(* IEC 61131-3 sources: 2026_Projet_YGO_ExcavatriceDragage/TOOLS/TEST_AUTO_CI/RESULTS/L_SIMULATION/tests (part 2) *)

TEST 'TC-T418-005 Perte permis stimulus et conflit en mouvement'
VAR
    fb : FB_Sim_Joystick;
    i : INT;
END_VAR
    fb.Enable := TRUE; fb(); fb.BtnRev_Down_Open := TRUE;
    ADVANCE_TIME(10000000); fb();
ADVANCE_TIME(10000000); fb();
ADVANCE_TIME(10000000); fb();
ADVANCE_TIME(10000000); fb();
ADVANCE_TIME(10000000); fb();
ADVANCE_TIME(10000000); fb();
ADVANCE_TIME(10000000); fb();
ADVANCE_TIME(10000000); fb();
ADVANCE_TIME(10000000); fb();
ADVANCE_TIME(10000000); fb();
ADVANCE_TIME(10000000); fb();
ADVANCE_TIME(10000000); fb();
ADVANCE_TIME(10000000); fb();
ADVANCE_TIME(10000000); fb();
ADVANCE_TIME(10000000); fb();
ADVANCE_TIME(10000000); fb();
ADVANCE_TIME(10000000); fb();
ADVANCE_TIME(10000000); fb();
ADVANCE_TIME(10000000); fb();
ADVANCE_TIME(10000000); fb();
ADVANCE_TIME(10000000); fb();
ADVANCE_TIME(10000000); fb();
ADVANCE_TIME(10000000); fb();
ADVANCE_TIME(10000000); fb();
ADVANCE_TIME(10000000); fb();
ADVANCE_TIME(10000000); fb();
ADVANCE_TIME(10000000); fb();
ADVANCE_TIME(10000000); fb();
ADVANCE_TIME(10000000); fb();
ADVANCE_TIME(10000000); fb();
ADVANCE_TIME(10000000); fb();
ADVANCE_TIME(10000000); fb();
ADVANCE_TIME(10000000); fb();
ADVANCE_TIME(10000000); fb();
ADVANCE_TIME(10000000); fb();
ADVANCE_TIME(10000000); fb();
ADVANCE_TIME(10000000); fb();
ADVANCE_TIME(10000000); fb();
ADVANCE_TIME(10000000); fb();
ADVANCE_TIME(10000000); fb();
ADVANCE_TIME(10000000); fb();
ADVANCE_TIME(10000000); fb();
ADVANCE_TIME(10000000); fb();
ADVANCE_TIME(10000000); fb();
ADVANCE_TIME(10000000); fb();
ADVANCE_TIME(10000000); fb();
ADVANCE_TIME(10000000); fb();
ADVANCE_TIME(10000000); fb();
ADVANCE_TIME(10000000); fb();
ADVANCE_TIME(10000000); fb();
ADVANCE_TIME(10000000); fb();
ADVANCE_TIME(10000000); fb();
ADVANCE_TIME(10000000); fb();
ADVANCE_TIME(10000000); fb();
ADVANCE_TIME(10000000); fb();
ADVANCE_TIME(10000000); fb();
ADVANCE_TIME(10000000); fb();
ADVANCE_TIME(10000000); fb();
ADVANCE_TIME(10000000); fb();
ADVANCE_TIME(10000000); fb();
ADVANCE_TIME(10000000); fb();
ADVANCE_TIME(10000000); fb();
ADVANCE_TIME(10000000); fb();
ADVANCE_TIME(10000000); fb();
ADVANCE_TIME(10000000); fb();
ADVANCE_TIME(10000000); fb();
ADVANCE_TIME(10000000); fb();
ADVANCE_TIME(10000000); fb();
ADVANCE_TIME(10000000); fb();
ADVANCE_TIME(10000000); fb();
ADVANCE_TIME(10000000); fb();
ADVANCE_TIME(10000000); fb();
ADVANCE_TIME(10000000); fb();
ADVANCE_TIME(10000000); fb();
ADVANCE_TIME(10000000); fb();
ADVANCE_TIME(10000000); fb();
ADVANCE_TIME(10000000); fb();
ADVANCE_TIME(10000000); fb();
ADVANCE_TIME(10000000); fb();
ADVANCE_TIME(10000000); fb();
ADVANCE_TIME(10000000); fb();
ADVANCE_TIME(10000000); fb();
ADVANCE_TIME(10000000); fb();
ADVANCE_TIME(10000000); fb();
ADVANCE_TIME(10000000); fb();
ADVANCE_TIME(10000000); fb();
ADVANCE_TIME(10000000); fb();
ADVANCE_TIME(10000000); fb();
ADVANCE_TIME(10000000); fb();
ADVANCE_TIME(10000000); fb();
ADVANCE_TIME(10000000); fb();
ADVANCE_TIME(10000000); fb();
ADVANCE_TIME(10000000); fb();
ADVANCE_TIME(10000000); fb();
ADVANCE_TIME(10000000); fb();
ADVANCE_TIME(10000000); fb();
ADVANCE_TIME(10000000); fb();
ADVANCE_TIME(10000000); fb();
ADVANCE_TIME(10000000); fb();
ADVANCE_TIME(10000000); fb();
    ASSERT_TRUE(fb.RawY < 5000, 'Y negatif');
    fb.GesturePermit := FALSE; fb();
    ASSERT_FALSE(fb.RawButton, 'Retrait permis simulateur annule bouton');
    fb.GesturePermit := TRUE;
    ADVANCE_TIME(10000000); fb();
        ASSERT_FALSE(fb.RawButton, 'Retour permis ne rearme pas');
ADVANCE_TIME(10000000); fb();
        ASSERT_FALSE(fb.RawButton, 'Retour permis ne rearme pas');
ADVANCE_TIME(10000000); fb();
        ASSERT_FALSE(fb.RawButton, 'Retour permis ne rearme pas');
ADVANCE_TIME(10000000); fb();
        ASSERT_FALSE(fb.RawButton, 'Retour permis ne rearme pas');
ADVANCE_TIME(10000000); fb();
        ASSERT_FALSE(fb.RawButton, 'Retour permis ne rearme pas');
ADVANCE_TIME(10000000); fb();
        ASSERT_FALSE(fb.RawButton, 'Retour permis ne rearme pas');
ADVANCE_TIME(10000000); fb();
        ASSERT_FALSE(fb.RawButton, 'Retour permis ne rearme pas');
ADVANCE_TIME(10000000); fb();
        ASSERT_FALSE(fb.RawButton, 'Retour permis ne rearme pas');
ADVANCE_TIME(10000000); fb();
        ASSERT_FALSE(fb.RawButton, 'Retour permis ne rearme pas');
ADVANCE_TIME(10000000); fb();
        ASSERT_FALSE(fb.RawButton, 'Retour permis ne rearme pas');
ADVANCE_TIME(10000000); fb();
        ASSERT_FALSE(fb.RawButton, 'Retour permis ne rearme pas');
ADVANCE_TIME(10000000); fb();
        ASSERT_FALSE(fb.RawButton, 'Retour permis ne rearme pas');
ADVANCE_TIME(10000000); fb();
        ASSERT_FALSE(fb.RawButton, 'Retour permis ne rearme pas');
ADVANCE_TIME(10000000); fb();
        ASSERT_FALSE(fb.RawButton, 'Retour permis ne rearme pas');
ADVANCE_TIME(10000000); fb();
        ASSERT_FALSE(fb.RawButton, 'Retour permis ne rearme pas');
ADVANCE_TIME(10000000); fb();
        ASSERT_FALSE(fb.RawButton, 'Retour permis ne rearme pas');
ADVANCE_TIME(10000000); fb();
        ASSERT_FALSE(fb.RawButton, 'Retour permis ne rearme pas');
ADVANCE_TIME(10000000); fb();
        ASSERT_FALSE(fb.RawButton, 'Retour permis ne rearme pas');
ADVANCE_TIME(10000000); fb();
        ASSERT_FALSE(fb.RawButton, 'Retour permis ne rearme pas');
ADVANCE_TIME(10000000); fb();
        ASSERT_FALSE(fb.RawButton, 'Retour permis ne rearme pas');
ADVANCE_TIME(10000000); fb();
        ASSERT_FALSE(fb.RawButton, 'Retour permis ne rearme pas');
ADVANCE_TIME(10000000); fb();
        ASSERT_FALSE(fb.RawButton, 'Retour permis ne rearme pas');
ADVANCE_TIME(10000000); fb();
        ASSERT_FALSE(fb.RawButton, 'Retour permis ne rearme pas');
ADVANCE_TIME(10000000); fb();
        ASSERT_FALSE(fb.RawButton, 'Retour permis ne rearme pas');
ADVANCE_TIME(10000000); fb();
        ASSERT_FALSE(fb.RawButton, 'Retour permis ne rearme pas');
ADVANCE_TIME(10000000); fb();
        ASSERT_FALSE(fb.RawButton, 'Retour permis ne rearme pas');
ADVANCE_TIME(10000000); fb();
        ASSERT_FALSE(fb.RawButton, 'Retour permis ne rearme pas');
ADVANCE_TIME(10000000); fb();
        ASSERT_FALSE(fb.RawButton, 'Retour permis ne rearme pas');
ADVANCE_TIME(10000000); fb();
        ASSERT_FALSE(fb.RawButton, 'Retour permis ne rearme pas');
ADVANCE_TIME(10000000); fb();
        ASSERT_FALSE(fb.RawButton, 'Retour permis ne rearme pas');
ADVANCE_TIME(10000000); fb();
        ASSERT_FALSE(fb.RawButton, 'Retour permis ne rearme pas');
ADVANCE_TIME(10000000); fb();
        ASSERT_FALSE(fb.RawButton, 'Retour permis ne rearme pas');
ADVANCE_TIME(10000000); fb();
        ASSERT_FALSE(fb.RawButton, 'Retour permis ne rearme pas');
ADVANCE_TIME(10000000); fb();
        ASSERT_FALSE(fb.RawButton, 'Retour permis ne rearme pas');
ADVANCE_TIME(10000000); fb();
        ASSERT_FALSE(fb.RawButton, 'Retour permis ne rearme pas');
ADVANCE_TIME(10000000); fb();
        ASSERT_FALSE(fb.RawButton, 'Retour permis ne rearme pas');
ADVANCE_TIME(10000000); fb();
        ASSERT_FALSE(fb.RawButton, 'Retour permis ne rearme pas');
ADVANCE_TIME(10000000); fb();
        ASSERT_FALSE(fb.RawButton, 'Retour permis ne rearme pas');
ADVANCE_TIME(10000000); fb();
        ASSERT_FALSE(fb.RawButton, 'Retour permis ne rearme pas');
ADVANCE_TIME(10000000); fb();
        ASSERT_FALSE(fb.RawButton, 'Retour permis ne rearme pas');
ADVANCE_TIME(10000000); fb();
        ASSERT_FALSE(fb.RawButton, 'Retour permis ne rearme pas');
ADVANCE_TIME(10000000); fb();
        ASSERT_FALSE(fb.RawButton, 'Retour permis ne rearme pas');
ADVANCE_TIME(10000000); fb();
        ASSERT_FALSE(fb.RawButton, 'Retour permis ne rearme pas');
ADVANCE_TIME(10000000); fb();
        ASSERT_FALSE(fb.RawButton, 'Retour permis ne rearme pas');
ADVANCE_TIME(10000000); fb();
        ASSERT_FALSE(fb.RawButton, 'Retour permis ne rearme pas');
ADVANCE_TIME(10000000); fb();
        ASSERT_FALSE(fb.RawButton, 'Retour permis ne rearme pas');
ADVANCE_TIME(10000000); fb();
        ASSERT_FALSE(fb.RawButton, 'Retour permis ne rearme pas');
ADVANCE_TIME(10000000); fb();
        ASSERT_FALSE(fb.RawButton, 'Retour permis ne rearme pas');
ADVANCE_TIME(10000000); fb();
        ASSERT_FALSE(fb.RawButton, 'Retour permis ne rearme pas');
ADVANCE_TIME(10000000); fb();
        ASSERT_FALSE(fb.RawButton, 'Retour permis ne rearme pas');
ADVANCE_TIME(10000000); fb();
        ASSERT_FALSE(fb.RawButton, 'Retour permis ne rearme pas');
ADVANCE_TIME(10000000); fb();
        ASSERT_FALSE(fb.RawButton, 'Retour permis ne rearme pas');
ADVANCE_TIME(10000000); fb();
        ASSERT_FALSE(fb.RawButton, 'Retour permis ne rearme pas');
ADVANCE_TIME(10000000); fb();
        ASSERT_FALSE(fb.RawButton, 'Retour permis ne rearme pas');
ADVANCE_TIME(10000000); fb();
        ASSERT_FALSE(fb.RawButton, 'Retour permis ne rearme pas');
ADVANCE_TIME(10000000); fb();
        ASSERT_FALSE(fb.RawButton, 'Retour permis ne rearme pas');
ADVANCE_TIME(10000000); fb();
        ASSERT_FALSE(fb.RawButton, 'Retour permis ne rearme pas');
ADVANCE_TIME(10000000); fb();
        ASSERT_FALSE(fb.RawButton, 'Retour permis ne rearme pas');
ADVANCE_TIME(10000000); fb();
        ASSERT_FALSE(fb.RawButton, 'Retour permis ne rearme pas');
ADVANCE_TIME(10000000); fb();
        ASSERT_FALSE(fb.RawButton, 'Retour permis ne rearme pas');
ADVANCE_TIME(10000000); fb();
        ASSERT_FALSE(fb.RawButton, 'Retour permis ne rearme pas');
ADVANCE_TIME(10000000); fb();
        ASSERT_FALSE(fb.RawButton, 'Retour permis ne rearme pas');
ADVANCE_TIME(10000000); fb();
        ASSERT_FALSE(fb.RawButton, 'Retour permis ne rearme pas');
ADVANCE_TIME(10000000); fb();
        ASSERT_FALSE(fb.RawButton, 'Retour permis ne rearme pas');
ADVANCE_TIME(10000000); fb();
        ASSERT_FALSE(fb.RawButton, 'Retour permis ne rearme pas');
ADVANCE_TIME(10000000); fb();
        ASSERT_FALSE(fb.RawButton, 'Retour permis ne rearme pas');
ADVANCE_TIME(10000000); fb();
        ASSERT_FALSE(fb.RawButton, 'Retour permis ne rearme pas');
ADVANCE_TIME(10000000); fb();
        ASSERT_FALSE(fb.RawButton, 'Retour permis ne rearme pas');
ADVANCE_TIME(10000000); fb();
        ASSERT_FALSE(fb.RawButton, 'Retour permis ne rearme pas');
ADVANCE_TIME(10000000); fb();
        ASSERT_FALSE(fb.RawButton, 'Retour permis ne rearme pas');
ADVANCE_TIME(10000000); fb();
        ASSERT_FALSE(fb.RawButton, 'Retour permis ne rearme pas');
ADVANCE_TIME(10000000); fb();
        ASSERT_FALSE(fb.RawButton, 'Retour permis ne rearme pas');
ADVANCE_TIME(10000000); fb();
        ASSERT_FALSE(fb.RawButton, 'Retour permis ne rearme pas');
ADVANCE_TIME(10000000); fb();
        ASSERT_FALSE(fb.RawButton, 'Retour permis ne rearme pas');
ADVANCE_TIME(10000000); fb();
        ASSERT_FALSE(fb.RawButton, 'Retour permis ne rearme pas');
ADVANCE_TIME(10000000); fb();
        ASSERT_FALSE(fb.RawButton, 'Retour permis ne rearme pas');
ADVANCE_TIME(10000000); fb();
        ASSERT_FALSE(fb.RawButton, 'Retour permis ne rearme pas');
ADVANCE_TIME(10000000); fb();
        ASSERT_FALSE(fb.RawButton, 'Retour permis ne rearme pas');
ADVANCE_TIME(10000000); fb();
        ASSERT_FALSE(fb.RawButton, 'Retour permis ne rearme pas');
ADVANCE_TIME(10000000); fb();
        ASSERT_FALSE(fb.RawButton, 'Retour permis ne rearme pas');
ADVANCE_TIME(10000000); fb();
        ASSERT_FALSE(fb.RawButton, 'Retour permis ne rearme pas');
ADVANCE_TIME(10000000); fb();
        ASSERT_FALSE(fb.RawButton, 'Retour permis ne rearme pas');
ADVANCE_TIME(10000000); fb();
        ASSERT_FALSE(fb.RawButton, 'Retour permis ne rearme pas');
ADVANCE_TIME(10000000); fb();
        ASSERT_FALSE(fb.RawButton, 'Retour permis ne rearme pas');
ADVANCE_TIME(10000000); fb();
        ASSERT_FALSE(fb.RawButton, 'Retour permis ne rearme pas');
ADVANCE_TIME(10000000); fb();
        ASSERT_FALSE(fb.RawButton, 'Retour permis ne rearme pas');
ADVANCE_TIME(10000000); fb();
        ASSERT_FALSE(fb.RawButton, 'Retour permis ne rearme pas');
ADVANCE_TIME(10000000); fb();
        ASSERT_FALSE(fb.RawButton, 'Retour permis ne rearme pas');
ADVANCE_TIME(10000000); fb();
        ASSERT_FALSE(fb.RawButton, 'Retour permis ne rearme pas');
ADVANCE_TIME(10000000); fb();
        ASSERT_FALSE(fb.RawButton, 'Retour permis ne rearme pas');
ADVANCE_TIME(10000000); fb();
        ASSERT_FALSE(fb.RawButton, 'Retour permis ne rearme pas');
ADVANCE_TIME(10000000); fb();
        ASSERT_FALSE(fb.RawButton, 'Retour permis ne rearme pas');
ADVANCE_TIME(10000000); fb();
        ASSERT_FALSE(fb.RawButton, 'Retour permis ne rearme pas');
ADVANCE_TIME(10000000); fb();
        ASSERT_FALSE(fb.RawButton, 'Retour permis ne rearme pas');
ADVANCE_TIME(10000000); fb();
        ASSERT_FALSE(fb.RawButton, 'Retour permis ne rearme pas');
ADVANCE_TIME(10000000); fb();
        ASSERT_FALSE(fb.RawButton, 'Retour permis ne rearme pas');
ADVANCE_TIME(10000000); fb();
        ASSERT_FALSE(fb.RawButton, 'Retour permis ne rearme pas');
ADVANCE_TIME(10000000); fb();
        ASSERT_FALSE(fb.RawButton, 'Retour permis ne rearme pas');
ADVANCE_TIME(10000000); fb();
        ASSERT_FALSE(fb.RawButton, 'Retour permis ne rearme pas');
ADVANCE_TIME(10000000); fb();
        ASSERT_FALSE(fb.RawButton, 'Retour permis ne rearme pas');
    ASSERT_EQ(fb.RawY, 5000, 'Retour neutre');
    fb.BtnRev_Down_Open := FALSE; fb(); fb.BtnFwd_Up_Close := TRUE;
    ADVANCE_TIME(10000000); fb();
ADVANCE_TIME(10000000); fb();
ADVANCE_TIME(10000000); fb();
ADVANCE_TIME(10000000); fb();
ADVANCE_TIME(10000000); fb();
ADVANCE_TIME(10000000); fb();
ADVANCE_TIME(10000000); fb();
ADVANCE_TIME(10000000); fb();
ADVANCE_TIME(10000000); fb();
ADVANCE_TIME(10000000); fb();
ADVANCE_TIME(10000000); fb();
ADVANCE_TIME(10000000); fb();
ADVANCE_TIME(10000000); fb();
ADVANCE_TIME(10000000); fb();
ADVANCE_TIME(10000000); fb();
ADVANCE_TIME(10000000); fb();
ADVANCE_TIME(10000000); fb();
ADVANCE_TIME(10000000); fb();
ADVANCE_TIME(10000000); fb();
ADVANCE_TIME(10000000); fb();
ADVANCE_TIME(10000000); fb();
ADVANCE_TIME(10000000); fb();
ADVANCE_TIME(10000000); fb();
ADVANCE_TIME(10000000); fb();
ADVANCE_TIME(10000000); fb();
ADVANCE_TIME(10000000); fb();
ADVANCE_TIME(10000000); fb();
ADVANCE_TIME(10000000); fb();
ADVANCE_TIME(10000000); fb();
ADVANCE_TIME(10000000); fb();
ADVANCE_TIME(10000000); fb();
ADVANCE_TIME(10000000); fb();
ADVANCE_TIME(10000000); fb();
ADVANCE_TIME(10000000); fb();
ADVANCE_TIME(10000000); fb();
ADVANCE_TIME(10000000); fb();
ADVANCE_TIME(10000000); fb();
ADVANCE_TIME(10000000); fb();
ADVANCE_TIME(10000000); fb();
ADVANCE_TIME(10000000); fb();
ADVANCE_TIME(10000000); fb();
ADVANCE_TIME(10000000); fb();
ADVANCE_TIME(10000000); fb();
ADVANCE_TIME(10000000); fb();
ADVANCE_TIME(10000000); fb();
ADVANCE_TIME(10000000); fb();
ADVANCE_TIME(10000000); fb();
ADVANCE_TIME(10000000); fb();
ADVANCE_TIME(10000000); fb();
ADVANCE_TIME(10000000); fb();
ADVANCE_TIME(10000000); fb();
ADVANCE_TIME(10000000); fb();
ADVANCE_TIME(10000000); fb();
ADVANCE_TIME(10000000); fb();
ADVANCE_TIME(10000000); fb();
ADVANCE_TIME(10000000); fb();
ADVANCE_TIME(10000000); fb();
ADVANCE_TIME(10000000); fb();
ADVANCE_TIME(10000000); fb();
ADVANCE_TIME(10000000); fb();
ADVANCE_TIME(10000000); fb();
ADVANCE_TIME(10000000); fb();
ADVANCE_TIME(10000000); fb();
ADVANCE_TIME(10000000); fb();
ADVANCE_TIME(10000000); fb();
ADVANCE_TIME(10000000); fb();
ADVANCE_TIME(10000000); fb();
ADVANCE_TIME(10000000); fb();
ADVANCE_TIME(10000000); fb();
ADVANCE_TIME(10000000); fb();
ADVANCE_TIME(10000000); fb();
ADVANCE_TIME(10000000); fb();
ADVANCE_TIME(10000000); fb();
ADVANCE_TIME(10000000); fb();
ADVANCE_TIME(10000000); fb();
ADVANCE_TIME(10000000); fb();
ADVANCE_TIME(10000000); fb();
ADVANCE_TIME(10000000); fb();
ADVANCE_TIME(10000000); fb();
ADVANCE_TIME(10000000); fb();
ADVANCE_TIME(10000000); fb();
ADVANCE_TIME(10000000); fb();
ADVANCE_TIME(10000000); fb();
ADVANCE_TIME(10000000); fb();
ADVANCE_TIME(10000000); fb();
ADVANCE_TIME(10000000); fb();
ADVANCE_TIME(10000000); fb();
ADVANCE_TIME(10000000); fb();
ADVANCE_TIME(10000000); fb();
ADVANCE_TIME(10000000); fb();
ADVANCE_TIME(10000000); fb();
ADVANCE_TIME(10000000); fb();
ADVANCE_TIME(10000000); fb();
ADVANCE_TIME(10000000); fb();
ADVANCE_TIME(10000000); fb();
ADVANCE_TIME(10000000); fb();
ADVANCE_TIME(10000000); fb();
ADVANCE_TIME(10000000); fb();
ADVANCE_TIME(10000000); fb();
ADVANCE_TIME(10000000); fb();
    fb.BtnRight_Fwd_MAINT := TRUE;
    ADVANCE_TIME(10000000); fb();
ADVANCE_TIME(10000000); fb();
ADVANCE_TIME(10000000); fb();
ADVANCE_TIME(10000000); fb();
ADVANCE_TIME(10000000); fb();
ADVANCE_TIME(10000000); fb();
ADVANCE_TIME(10000000); fb();
ADVANCE_TIME(10000000); fb();
ADVANCE_TIME(10000000); fb();
ADVANCE_TIME(10000000); fb();
ADVANCE_TIME(10000000); fb();
ADVANCE_TIME(10000000); fb();
ADVANCE_TIME(10000000); fb();
ADVANCE_TIME(10000000); fb();
ADVANCE_TIME(10000000); fb();
ADVANCE_TIME(10000000); fb();
ADVANCE_TIME(10000000); fb();
ADVANCE_TIME(10000000); fb();
ADVANCE_TIME(10000000); fb();
ADVANCE_TIME(10000000); fb();
ADVANCE_TIME(10000000); fb();
ADVANCE_TIME(10000000); fb();
ADVANCE_TIME(10000000); fb();
ADVANCE_TIME(10000000); fb();
ADVANCE_TIME(10000000); fb();
ADVANCE_TIME(10000000); fb();
ADVANCE_TIME(10000000); fb();
ADVANCE_TIME(10000000); fb();
ADVANCE_TIME(10000000); fb();
ADVANCE_TIME(10000000); fb();
ADVANCE_TIME(10000000); fb();
ADVANCE_TIME(10000000); fb();
ADVANCE_TIME(10000000); fb();
ADVANCE_TIME(10000000); fb();
ADVANCE_TIME(10000000); fb();
ADVANCE_TIME(10000000); fb();
ADVANCE_TIME(10000000); fb();
ADVANCE_TIME(10000000); fb();
ADVANCE_TIME(10000000); fb();
ADVANCE_TIME(10000000); fb();
ADVANCE_TIME(10000000); fb();
ADVANCE_TIME(10000000); fb();
ADVANCE_TIME(10000000); fb();
ADVANCE_TIME(10000000); fb();
ADVANCE_TIME(10000000); fb();
ADVANCE_TIME(10000000); fb();
ADVANCE_TIME(10000000); fb();
ADVANCE_TIME(10000000); fb();
ADVANCE_TIME(10000000); fb();
ADVANCE_TIME(10000000); fb();
ADVANCE_TIME(10000000); fb();
ADVANCE_TIME(10000000); fb();
ADVANCE_TIME(10000000); fb();
ADVANCE_TIME(10000000); fb();
ADVANCE_TIME(10000000); fb();
ADVANCE_TIME(10000000); fb();
ADVANCE_TIME(10000000); fb();
ADVANCE_TIME(10000000); fb();
ADVANCE_TIME(10000000); fb();
ADVANCE_TIME(10000000); fb();
ADVANCE_TIME(10000000); fb();
ADVANCE_TIME(10000000); fb();
ADVANCE_TIME(10000000); fb();
ADVANCE_TIME(10000000); fb();
ADVANCE_TIME(10000000); fb();
ADVANCE_TIME(10000000); fb();
ADVANCE_TIME(10000000); fb();
ADVANCE_TIME(10000000); fb();
ADVANCE_TIME(10000000); fb();
ADVANCE_TIME(10000000); fb();
ADVANCE_TIME(10000000); fb();
ADVANCE_TIME(10000000); fb();
ADVANCE_TIME(10000000); fb();
ADVANCE_TIME(10000000); fb();
ADVANCE_TIME(10000000); fb();
ADVANCE_TIME(10000000); fb();
ADVANCE_TIME(10000000); fb();
ADVANCE_TIME(10000000); fb();
ADVANCE_TIME(10000000); fb();
ADVANCE_TIME(10000000); fb();
ADVANCE_TIME(10000000); fb();
ADVANCE_TIME(10000000); fb();
ADVANCE_TIME(10000000); fb();
ADVANCE_TIME(10000000); fb();
ADVANCE_TIME(10000000); fb();
ADVANCE_TIME(10000000); fb();
ADVANCE_TIME(10000000); fb();
ADVANCE_TIME(10000000); fb();
ADVANCE_TIME(10000000); fb();
ADVANCE_TIME(10000000); fb();
ADVANCE_TIME(10000000); fb();
ADVANCE_TIME(10000000); fb();
ADVANCE_TIME(10000000); fb();
ADVANCE_TIME(10000000); fb();
ADVANCE_TIME(10000000); fb();
ADVANCE_TIME(10000000); fb();
ADVANCE_TIME(10000000); fb();
ADVANCE_TIME(10000000); fb();
ADVANCE_TIME(10000000); fb();
ADVANCE_TIME(10000000); fb();
    ASSERT_EQ(fb.RawY, 5000, 'Conflit en mouvement retourne au neutre');
    ASSERT_FALSE(fb.RawButton, 'Conflit ne produit pas appui');
END_TEST

TEST 'TC-T418-006 Dynamiques depassement et bagotement conservees'
VAR
    fb : FB_Sim_Joystick;
    i : INT;
    oscillationSeen : BOOL;
END_VAR
    oscillationSeen := FALSE;
    fb.Enable := TRUE; fb.OvershootActive := TRUE; fb.BagotementActive := TRUE;
    fb(); fb.BtnRight_Fwd_MAINT := TRUE;
    ADVANCE_TIME(10000000); fb();
ADVANCE_TIME(10000000); fb();
ADVANCE_TIME(10000000); fb();
ADVANCE_TIME(10000000); fb();
ADVANCE_TIME(10000000); fb();
ADVANCE_TIME(10000000); fb();
ADVANCE_TIME(10000000); fb();
ADVANCE_TIME(10000000); fb();
ADVANCE_TIME(10000000); fb();
ADVANCE_TIME(10000000); fb();
ADVANCE_TIME(10000000); fb();
ADVANCE_TIME(10000000); fb();
ADVANCE_TIME(10000000); fb();
ADVANCE_TIME(10000000); fb();
ADVANCE_TIME(10000000); fb();
ADVANCE_TIME(10000000); fb();
ADVANCE_TIME(10000000); fb();
ADVANCE_TIME(10000000); fb();
ADVANCE_TIME(10000000); fb();
ADVANCE_TIME(10000000); fb();
ADVANCE_TIME(10000000); fb();
ADVANCE_TIME(10000000); fb();
ADVANCE_TIME(10000000); fb();
ADVANCE_TIME(10000000); fb();
ADVANCE_TIME(10000000); fb();
ADVANCE_TIME(10000000); fb();
ADVANCE_TIME(10000000); fb();
ADVANCE_TIME(10000000); fb();
ADVANCE_TIME(10000000); fb();
ADVANCE_TIME(10000000); fb();
ADVANCE_TIME(10000000); fb();
ADVANCE_TIME(10000000); fb();
ADVANCE_TIME(10000000); fb();
ADVANCE_TIME(10000000); fb();
ADVANCE_TIME(10000000); fb();
ADVANCE_TIME(10000000); fb();
ADVANCE_TIME(10000000); fb();
ADVANCE_TIME(10000000); fb();
ADVANCE_TIME(10000000); fb();
ADVANCE_TIME(10000000); fb();
ADVANCE_TIME(10000000); fb();
ADVANCE_TIME(10000000); fb();
ADVANCE_TIME(10000000); fb();
ADVANCE_TIME(10000000); fb();
ADVANCE_TIME(10000000); fb();
ADVANCE_TIME(10000000); fb();
ADVANCE_TIME(10000000); fb();
ADVANCE_TIME(10000000); fb();
ADVANCE_TIME(10000000); fb();
ADVANCE_TIME(10000000); fb();
ADVANCE_TIME(10000000); fb();
ADVANCE_TIME(10000000); fb();
ADVANCE_TIME(10000000); fb();
ADVANCE_TIME(10000000); fb();
ADVANCE_TIME(10000000); fb();
ADVANCE_TIME(10000000); fb();
ADVANCE_TIME(10000000); fb();
ADVANCE_TIME(10000000); fb();
ADVANCE_TIME(10000000); fb();
ADVANCE_TIME(10000000); fb();
ADVANCE_TIME(10000000); fb();
ADVANCE_TIME(10000000); fb();
ADVANCE_TIME(10000000); fb();
ADVANCE_TIME(10000000); fb();
ADVANCE_TIME(10000000); fb();
ADVANCE_TIME(10000000); fb();
ADVANCE_TIME(10000000); fb();
ADVANCE_TIME(10000000); fb();
ADVANCE_TIME(10000000); fb();
ADVANCE_TIME(10000000); fb();
ADVANCE_TIME(10000000); fb();
ADVANCE_TIME(10000000); fb();
ADVANCE_TIME(10000000); fb();
ADVANCE_TIME(10000000); fb();
ADVANCE_TIME(10000000); fb();
ADVANCE_TIME(10000000); fb();
ADVANCE_TIME(10000000); fb();
ADVANCE_TIME(10000000); fb();
ADVANCE_TIME(10000000); fb();
ADVANCE_TIME(10000000); fb();
ADVANCE_TIME(10000000); fb();
ADVANCE_TIME(10000000); fb();
ADVANCE_TIME(10000000); fb();
ADVANCE_TIME(10000000); fb();
ADVANCE_TIME(10000000); fb();
ADVANCE_TIME(10000000); fb();
ADVANCE_TIME(10000000); fb();
ADVANCE_TIME(10000000); fb();
ADVANCE_TIME(10000000); fb();
ADVANCE_TIME(10000000); fb();
ADVANCE_TIME(10000000); fb();
ADVANCE_TIME(10000000); fb();
ADVANCE_TIME(10000000); fb();
ADVANCE_TIME(10000000); fb();
ADVANCE_TIME(10000000); fb();
ADVANCE_TIME(10000000); fb();
ADVANCE_TIME(10000000); fb();
ADVANCE_TIME(10000000); fb();
ADVANCE_TIME(10000000); fb();
ADVANCE_TIME(10000000); fb();
ADVANCE_TIME(10000000); fb();
ADVANCE_TIME(10000000); fb();
ADVANCE_TIME(10000000); fb();
ADVANCE_TIME(10000000); fb();
ADVANCE_TIME(10000000); fb();
ADVANCE_TIME(10000000); fb();
ADVANCE_TIME(10000000); fb();
ADVANCE_TIME(10000000); fb();
ADVANCE_TIME(10000000); fb();
ADVANCE_TIME(10000000); fb();
ADVANCE_TIME(10000000); fb();
ADVANCE_TIME(10000000); fb();
ADVANCE_TIME(10000000); fb();
ADVANCE_TIME(10000000); fb();
ADVANCE_TIME(10000000); fb();
ADVANCE_TIME(10000000); fb();
ADVANCE_TIME(10000000); fb();
ADVANCE_TIME(10000000); fb();
ADVANCE_TIME(10000000); fb();
ADVANCE_TIME(10000000); fb();
ADVANCE_TIME(10000000); fb();
ADVANCE_TIME(10000000); fb();
ADVANCE_TIME(10000000); fb();
ADVANCE_TIME(10000000); fb();
ADVANCE_TIME(10000000); fb();
ADVANCE_TIME(10000000); fb();
ADVANCE_TIME(10000000); fb();
ADVANCE_TIME(10000000); fb();
ADVANCE_TIME(10000000); fb();
ADVANCE_TIME(10000000); fb();
ADVANCE_TIME(10000000); fb();
ADVANCE_TIME(10000000); fb();
ADVANCE_TIME(10000000); fb();
ADVANCE_TIME(10000000); fb();
ADVANCE_TIME(10000000); fb();
ADVANCE_TIME(10000000); fb();
ADVANCE_TIME(10000000); fb();
ADVANCE_TIME(10000000); fb();
ADVANCE_TIME(10000000); fb();
ADVANCE_TIME(10000000); fb();
ADVANCE_TIME(10000000); fb();
ADVANCE_TIME(10000000); fb();
ADVANCE_TIME(10000000); fb();
ADVANCE_TIME(10000000); fb();
ADVANCE_TIME(10000000); fb();
ADVANCE_TIME(10000000); fb();
ADVANCE_TIME(10000000); fb();
ADVANCE_TIME(10000000); fb();
ADVANCE_TIME(10000000); fb();
ADVANCE_TIME(10000000); fb();
ADVANCE_TIME(10000000); fb();
ADVANCE_TIME(10000000); fb();
ADVANCE_TIME(10000000); fb();
ADVANCE_TIME(10000000); fb();
ADVANCE_TIME(10000000); fb();
ADVANCE_TIME(10000000); fb();
ADVANCE_TIME(10000000); fb();
ADVANCE_TIME(10000000); fb();
ADVANCE_TIME(10000000); fb();
ADVANCE_TIME(10000000); fb();
ADVANCE_TIME(10000000); fb();
ADVANCE_TIME(10000000); fb();
ADVANCE_TIME(10000000); fb();
ADVANCE_TIME(10000000); fb();
ADVANCE_TIME(10000000); fb();
ADVANCE_TIME(10000000); fb();
ADVANCE_TIME(10000000); fb();
ADVANCE_TIME(10000000); fb();
ADVANCE_TIME(10000000); fb();
ADVANCE_TIME(10000000); fb();
ADVANCE_TIME(10000000); fb();
ADVANCE_TIME(10000000); fb();
ADVANCE_TIME(10000000); fb();
ADVANCE_TIME(10000000); fb();
ADVANCE_TIME(10000000); fb();
ADVANCE_TIME(10000000); fb();
ADVANCE_TIME(10000000); fb();
ADVANCE_TIME(10000000); fb();
ADVANCE_TIME(10000000); fb();
ADVANCE_TIME(10000000); fb();
ADVANCE_TIME(10000000); fb();
ADVANCE_TIME(10000000); fb();
ADVANCE_TIME(10000000); fb();
ADVANCE_TIME(10000000); fb();
ADVANCE_TIME(10000000); fb();
ADVANCE_TIME(10000000); fb();
ADVANCE_TIME(10000000); fb();
ADVANCE_TIME(10000000); fb();
ADVANCE_TIME(10000000); fb();
ADVANCE_TIME(10000000); fb();
ADVANCE_TIME(10000000); fb();
ADVANCE_TIME(10000000); fb();
ADVANCE_TIME(10000000); fb();
ADVANCE_TIME(10000000); fb();
ADVANCE_TIME(10000000); fb();
ADVANCE_TIME(10000000); fb();
ADVANCE_TIME(10000000); fb();
ADVANCE_TIME(10000000); fb();
ADVANCE_TIME(10000000); fb();
ADVANCE_TIME(10000000); fb();
ADVANCE_TIME(10000000); fb();
ADVANCE_TIME(10000000); fb();
ADVANCE_TIME(10000000); fb();
ADVANCE_TIME(10000000); fb();
ADVANCE_TIME(10000000); fb();
ADVANCE_TIME(10000000); fb();
ADVANCE_TIME(10000000); fb();
ADVANCE_TIME(10000000); fb();
ADVANCE_TIME(10000000); fb();
ADVANCE_TIME(10000000); fb();
ADVANCE_TIME(10000000); fb();
ADVANCE_TIME(10000000); fb();
ADVANCE_TIME(10000000); fb();
ADVANCE_TIME(10000000); fb();
ADVANCE_TIME(10000000); fb();
ADVANCE_TIME(10000000); fb();
ADVANCE_TIME(10000000); fb();
ADVANCE_TIME(10000000); fb();
ADVANCE_TIME(10000000); fb();
ADVANCE_TIME(10000000); fb();
ADVANCE_TIME(10000000); fb();
ADVANCE_TIME(10000000); fb();
ADVANCE_TIME(10000000); fb();
ADVANCE_TIME(10000000); fb();
ADVANCE_TIME(10000000); fb();
ADVANCE_TIME(10000000); fb();
ADVANCE_TIME(10000000); fb();
ADVANCE_TIME(10000000); fb();
ADVANCE_TIME(10000000); fb();
ADVANCE_TIME(10000000); fb();
ADVANCE_TIME(10000000); fb();
ADVANCE_TIME(10000000); fb();
ADVANCE_TIME(10000000); fb();
ADVANCE_TIME(10000000); fb();
ADVANCE_TIME(10000000); fb();
ADVANCE_TIME(10000000); fb();
ADVANCE_TIME(10000000); fb();
ADVANCE_TIME(10000000); fb();
ADVANCE_TIME(10000000); fb();
ADVANCE_TIME(10000000); fb();
ADVANCE_TIME(10000000); fb();
ADVANCE_TIME(10000000); fb();
ADVANCE_TIME(10000000); fb();
ADVANCE_TIME(10000000); fb();
ADVANCE_TIME(10000000); fb();
ADVANCE_TIME(10000000); fb();
ADVANCE_TIME(10000000); fb();
ADVANCE_TIME(10000000); fb();
ADVANCE_TIME(10000000); fb();
ADVANCE_TIME(10000000); fb();
    ASSERT_TRUE(fb.RawX > 10500, 'Injection depassement capteur conservee');
    fb.BtnRight_Fwd_MAINT := FALSE;
    ADVANCE_TIME(10000000); fb();
        IF fb.RawX < 5000 THEN oscillationSeen := TRUE; END_IF;
        ASSERT_FALSE(fb.RawButton, 'Aucun front pendant bagotement');
ADVANCE_TIME(10000000); fb();
        IF fb.RawX < 5000 THEN oscillationSeen := TRUE; END_IF;
        ASSERT_FALSE(fb.RawButton, 'Aucun front pendant bagotement');
ADVANCE_TIME(10000000); fb();
        IF fb.RawX < 5000 THEN oscillationSeen := TRUE; END_IF;
        ASSERT_FALSE(fb.RawButton, 'Aucun front pendant bagotement');
ADVANCE_TIME(10000000); fb();
        IF fb.RawX < 5000 THEN oscillationSeen := TRUE; END_IF;
        ASSERT_FALSE(fb.RawButton, 'Aucun front pendant bagotement');
ADVANCE_TIME(10000000); fb();
        IF fb.RawX < 5000 THEN oscillationSeen := TRUE; END_IF;
        ASSERT_FALSE(fb.RawButton, 'Aucun front pendant bagotement');
ADVANCE_TIME(10000000); fb();
        IF fb.RawX < 5000 THEN oscillationSeen := TRUE; END_IF;
        ASSERT_FALSE(fb.RawButton, 'Aucun front pendant bagotement');
ADVANCE_TIME(10000000); fb();
        IF fb.RawX < 5000 THEN oscillationSeen := TRUE; END_IF;
        ASSERT_FALSE(fb.RawButton, 'Aucun front pendant bagotement');
ADVANCE_TIME(10000000); fb();
        IF fb.RawX < 5000 THEN oscillationSeen := TRUE; END_IF;
        ASSERT_FALSE(fb.RawButton, 'Aucun front pendant bagotement');
ADVANCE_TIME(10000000); fb();
        IF fb.RawX < 5000 THEN oscillationSeen := TRUE; END_IF;
        ASSERT_FALSE(fb.RawButton, 'Aucun front pendant bagotement');
ADVANCE_TIME(10000000); fb();
        IF fb.RawX < 5000 THEN oscillationSeen := TRUE; END_IF;
        ASSERT_FALSE(fb.RawButton, 'Aucun front pendant bagotement');
ADVANCE_TIME(10000000); fb();
        IF fb.RawX < 5000 THEN oscillationSeen := TRUE; END_IF;
        ASSERT_FALSE(fb.RawButton, 'Aucun front pendant bagotement');
ADVANCE_TIME(10000000); fb();
        IF fb.RawX < 5000 THEN oscillationSeen := TRUE; END_IF;
        ASSERT_FALSE(fb.RawButton, 'Aucun front pendant bagotement');
ADVANCE_TIME(10000000); fb();
        IF fb.RawX < 5000 THEN oscillationSeen := TRUE; END_IF;
        ASSERT_FALSE(fb.RawButton, 'Aucun front pendant bagotement');
ADVANCE_TIME(10000000); fb();
        IF fb.RawX < 5000 THEN oscillationSeen := TRUE; END_IF;
        ASSERT_FALSE(fb.RawButton, 'Aucun front pendant bagotement');
ADVANCE_TIME(10000000); fb();
        IF fb.RawX < 5000 THEN oscillationSeen := TRUE; END_IF;
        ASSERT_FALSE(fb.RawButton, 'Aucun front pendant bagotement');
ADVANCE_TIME(10000000); fb();
        IF fb.RawX < 5000 THEN oscillationSeen := TRUE; END_IF;
        ASSERT_FALSE(fb.RawButton, 'Aucun front pendant bagotement');
ADVANCE_TIME(10000000); fb();
        IF fb.RawX < 5000 THEN oscillationSeen := TRUE; END_IF;
        ASSERT_FALSE(fb.RawButton, 'Aucun front pendant bagotement');
ADVANCE_TIME(10000000); fb();
        IF fb.RawX < 5000 THEN oscillationSeen := TRUE; END_IF;
        ASSERT_FALSE(fb.RawButton, 'Aucun front pendant bagotement');
ADVANCE_TIME(10000000); fb();
        IF fb.RawX < 5000 THEN oscillationSeen := TRUE; END_IF;
        ASSERT_FALSE(fb.RawButton, 'Aucun front pendant bagotement');
ADVANCE_TIME(10000000); fb();
        IF fb.RawX < 5000 THEN oscillationSeen := TRUE; END_IF;
        ASSERT_FALSE(fb.RawButton, 'Aucun front pendant bagotement');
ADVANCE_TIME(10000000); fb();
        IF fb.RawX < 5000 THEN oscillationSeen := TRUE; END_IF;
        ASSERT_FALSE(fb.RawButton, 'Aucun front pendant bagotement');
ADVANCE_TIME(10000000); fb();
        IF fb.RawX < 5000 THEN oscillationSeen := TRUE; END_IF;
        ASSERT_FALSE(fb.RawButton, 'Aucun front pendant bagotement');
ADVANCE_TIME(10000000); fb();
        IF fb.RawX < 5000 THEN oscillationSeen := TRUE; END_IF;
        ASSERT_FALSE(fb.RawButton, 'Aucun front pendant bagotement');
ADVANCE_TIME(10000000); fb();
        IF fb.RawX < 5000 THEN oscillationSeen := TRUE; END_IF;
        ASSERT_FALSE(fb.RawButton, 'Aucun front pendant bagotement');
ADVANCE_TIME(10000000); fb();
        IF fb.RawX < 5000 THEN oscillationSeen := TRUE; END_IF;
        ASSERT_FALSE(fb.RawButton, 'Aucun front pendant bagotement');
ADVANCE_TIME(10000000); fb();
        IF fb.RawX < 5000 THEN oscillationSeen := TRUE; END_IF;
        ASSERT_FALSE(fb.RawButton, 'Aucun front pendant bagotement');
ADVANCE_TIME(10000000); fb();
        IF fb.RawX < 5000 THEN oscillationSeen := TRUE; END_IF;
        ASSERT_FALSE(fb.RawButton, 'Aucun front pendant bagotement');
ADVANCE_TIME(10000000); fb();
        IF fb.RawX < 5000 THEN oscillationSeen := TRUE; END_IF;
        ASSERT_FALSE(fb.RawButton, 'Aucun front pendant bagotement');
ADVANCE_TIME(10000000); fb();
        IF fb.RawX < 5000 THEN oscillationSeen := TRUE; END_IF;
        ASSERT_FALSE(fb.RawButton, 'Aucun front pendant bagotement');
ADVANCE_TIME(10000000); fb();
        IF fb.RawX < 5000 THEN oscillationSeen := TRUE; END_IF;
        ASSERT_FALSE(fb.RawButton, 'Aucun front pendant bagotement');
ADVANCE_TIME(10000000); fb();
        IF fb.RawX < 5000 THEN oscillationSeen := TRUE; END_IF;
        ASSERT_FALSE(fb.RawButton, 'Aucun front pendant bagotement');
ADVANCE_TIME(10000000); fb();
        IF fb.RawX < 5000 THEN oscillationSeen := TRUE; END_IF;
        ASSERT_FALSE(fb.RawButton, 'Aucun front pendant bagotement');
ADVANCE_TIME(10000000); fb();
        IF fb.RawX < 5000 THEN oscillationSeen := TRUE; END_IF;
        ASSERT_FALSE(fb.RawButton, 'Aucun front pendant bagotement');
ADVANCE_TIME(10000000); fb();
        IF fb.RawX < 5000 THEN oscillationSeen := TRUE; END_IF;
        ASSERT_FALSE(fb.RawButton, 'Aucun front pendant bagotement');
ADVANCE_TIME(10000000); fb();
        IF fb.RawX < 5000 THEN oscillationSeen := TRUE; END_IF;
        ASSERT_FALSE(fb.RawButton, 'Aucun front pendant bagotement');
ADVANCE_TIME(10000000); fb();
        IF fb.RawX < 5000 THEN oscillationSeen := TRUE; END_IF;
        ASSERT_FALSE(fb.RawButton, 'Aucun front pendant bagotement');
ADVANCE_TIME(10000000); fb();
        IF fb.RawX < 5000 THEN oscillationSeen := TRUE; END_IF;
        ASSERT_FALSE(fb.RawButton, 'Aucun front pendant bagotement');
ADVANCE_TIME(10000000); fb();
        IF fb.RawX < 5000 THEN oscillationSeen := TRUE; END_IF;
        ASSERT_FALSE(fb.RawButton, 'Aucun front pendant bagotement');
ADVANCE_TIME(10000000); fb();
        IF fb.RawX < 5000 THEN oscillationSeen := TRUE; END_IF;
        ASSERT_FALSE(fb.RawButton, 'Aucun front pendant bagotement');
ADVANCE_TIME(10000000); fb();
        IF fb.RawX < 5000 THEN oscillationSeen := TRUE; END_IF;
        ASSERT_FALSE(fb.RawButton, 'Aucun front pendant bagotement');
ADVANCE_TIME(10000000); fb();
        IF fb.RawX < 5000 THEN oscillationSeen := TRUE; END_IF;
        ASSERT_FALSE(fb.RawButton, 'Aucun front pendant bagotement');
ADVANCE_TIME(10000000); fb();
        IF fb.RawX < 5000 THEN oscillationSeen := TRUE; END_IF;
        ASSERT_FALSE(fb.RawButton, 'Aucun front pendant bagotement');
ADVANCE_TIME(10000000); fb();
        IF fb.RawX < 5000 THEN oscillationSeen := TRUE; END_IF;
        ASSERT_FALSE(fb.RawButton, 'Aucun front pendant bagotement');
ADVANCE_TIME(10000000); fb();
        IF fb.RawX < 5000 THEN oscillationSeen := TRUE; END_IF;
        ASSERT_FALSE(fb.RawButton, 'Aucun front pendant bagotement');
ADVANCE_TIME(10000000); fb();
        IF fb.RawX < 5000 THEN oscillationSeen := TRUE; END_IF;
        ASSERT_FALSE(fb.RawButton, 'Aucun front pendant bagotement');
ADVANCE_TIME(10000000); fb();
        IF fb.RawX < 5000 THEN oscillationSeen := TRUE; END_IF;
        ASSERT_FALSE(fb.RawButton, 'Aucun front pendant bagotement');
ADVANCE_TIME(10000000); fb();
        IF fb.RawX < 5000 THEN oscillationSeen := TRUE; END_IF;
        ASSERT_FALSE(fb.RawButton, 'Aucun front pendant bagotement');
ADVANCE_TIME(10000000); fb();
        IF fb.RawX < 5000 THEN oscillationSeen := TRUE; END_IF;
        ASSERT_FALSE(fb.RawButton, 'Aucun front pendant bagotement');
ADVANCE_TIME(10000000); fb();
        IF fb.RawX < 5000 THEN oscillationSeen := TRUE; END_IF;
        ASSERT_FALSE(fb.RawButton, 'Aucun front pendant bagotement');
ADVANCE_TIME(10000000); fb();
        IF fb.RawX < 5000 THEN oscillationSeen := TRUE; END_IF;
        ASSERT_FALSE(fb.RawButton, 'Aucun front pendant bagotement');
ADVANCE_TIME(10000000); fb();
        IF fb.RawX < 5000 THEN oscillationSeen := TRUE; END_IF;
        ASSERT_FALSE(fb.RawButton, 'Aucun front pendant bagotement');
ADVANCE_TIME(10000000); fb();
        IF fb.RawX < 5000 THEN oscillationSeen := TRUE; END_IF;
        ASSERT_FALSE(fb.RawButton, 'Aucun front pendant bagotement');
ADVANCE_TIME(10000000); fb();
        IF fb.RawX < 5000 THEN oscillationSeen := TRUE; END_IF;
        ASSERT_FALSE(fb.RawButton, 'Aucun front pendant bagotement');
ADVANCE_TIME(10000000); fb();
        IF fb.RawX < 5000 THEN oscillationSeen := TRUE; END_IF;
        ASSERT_FALSE(fb.RawButton, 'Aucun front pendant bagotement');
ADVANCE_TIME(10000000); fb();
        IF fb.RawX < 5000 THEN oscillationSeen := TRUE; END_IF;
        ASSERT_FALSE(fb.RawButton, 'Aucun front pendant bagotement');
ADVANCE_TIME(10000000); fb();
        IF fb.RawX < 5000 THEN oscillationSeen := TRUE; END_IF;
        ASSERT_FALSE(fb.RawButton, 'Aucun front pendant bagotement');
ADVANCE_TIME(10000000); fb();
        IF fb.RawX < 5000 THEN oscillationSeen := TRUE; END_IF;
        ASSERT_FALSE(fb.RawButton, 'Aucun front pendant bagotement');
ADVANCE_TIME(10000000); fb();
        IF fb.RawX < 5000 THEN oscillationSeen := TRUE; END_IF;
        ASSERT_FALSE(fb.RawButton, 'Aucun front pendant bagotement');
ADVANCE_TIME(10000000); fb();
        IF fb.RawX < 5000 THEN oscillationSeen := TRUE; END_IF;
        ASSERT_FALSE(fb.RawButton, 'Aucun front pendant bagotement');
ADVANCE_TIME(10000000); fb();
        IF fb.RawX < 5000 THEN oscillationSeen := TRUE; END_IF;
        ASSERT_FALSE(fb.RawButton, 'Aucun front pendant bagotement');
ADVANCE_TIME(10000000); fb();
        IF fb.RawX < 5000 THEN oscillationSeen := TRUE; END_IF;
        ASSERT_FALSE(fb.RawButton, 'Aucun front pendant bagotement');
ADVANCE_TIME(10000000); fb();
        IF fb.RawX < 5000 THEN oscillationSeen := TRUE; END_IF;
        ASSERT_FALSE(fb.RawButton, 'Aucun front pendant bagotement');
ADVANCE_TIME(10000000); fb();
        IF fb.RawX < 5000 THEN oscillationSeen := TRUE; END_IF;
        ASSERT_FALSE(fb.RawButton, 'Aucun front pendant bagotement');
ADVANCE_TIME(10000000); fb();
        IF fb.RawX < 5000 THEN oscillationSeen := TRUE; END_IF;
        ASSERT_FALSE(fb.RawButton, 'Aucun front pendant bagotement');
ADVANCE_TIME(10000000); fb();
        IF fb.RawX < 5000 THEN oscillationSeen := TRUE; END_IF;
        ASSERT_FALSE(fb.RawButton, 'Aucun front pendant bagotement');
ADVANCE_TIME(10000000); fb();
        IF fb.RawX < 5000 THEN oscillationSeen := TRUE; END_IF;
        ASSERT_FALSE(fb.RawButton, 'Aucun front pendant bagotement');
ADVANCE_TIME(10000000); fb();
        IF fb.RawX < 5000 THEN oscillationSeen := TRUE; END_IF;
        ASSERT_FALSE(fb.RawButton, 'Aucun front pendant bagotement');
ADVANCE_TIME(10000000); fb();
        IF fb.RawX < 5000 THEN oscillationSeen := TRUE; END_IF;
        ASSERT_FALSE(fb.RawButton, 'Aucun front pendant bagotement');
ADVANCE_TIME(10000000); fb();
        IF fb.RawX < 5000 THEN oscillationSeen := TRUE; END_IF;
        ASSERT_FALSE(fb.RawButton, 'Aucun front pendant bagotement');
ADVANCE_TIME(10000000); fb();
        IF fb.RawX < 5000 THEN oscillationSeen := TRUE; END_IF;
        ASSERT_FALSE(fb.RawButton, 'Aucun front pendant bagotement');
ADVANCE_TIME(10000000); fb();
        IF fb.RawX < 5000 THEN oscillationSeen := TRUE; END_IF;
        ASSERT_FALSE(fb.RawButton, 'Aucun front pendant bagotement');
ADVANCE_TIME(10000000); fb();
        IF fb.RawX < 5000 THEN oscillationSeen := TRUE; END_IF;
        ASSERT_FALSE(fb.RawButton, 'Aucun front pendant bagotement');
ADVANCE_TIME(10000000); fb();
        IF fb.RawX < 5000 THEN oscillationSeen := TRUE; END_IF;
        ASSERT_FALSE(fb.RawButton, 'Aucun front pendant bagotement');
ADVANCE_TIME(10000000); fb();
        IF fb.RawX < 5000 THEN oscillationSeen := TRUE; END_IF;
        ASSERT_FALSE(fb.RawButton, 'Aucun front pendant bagotement');
ADVANCE_TIME(10000000); fb();
        IF fb.RawX < 5000 THEN oscillationSeen := TRUE; END_IF;
        ASSERT_FALSE(fb.RawButton, 'Aucun front pendant bagotement');
ADVANCE_TIME(10000000); fb();
        IF fb.RawX < 5000 THEN oscillationSeen := TRUE; END_IF;
        ASSERT_FALSE(fb.RawButton, 'Aucun front pendant bagotement');
ADVANCE_TIME(10000000); fb();
        IF fb.RawX < 5000 THEN oscillationSeen := TRUE; END_IF;
        ASSERT_FALSE(fb.RawButton, 'Aucun front pendant bagotement');
ADVANCE_TIME(10000000); fb();
        IF fb.RawX < 5000 THEN oscillationSeen := TRUE; END_IF;
        ASSERT_FALSE(fb.RawButton, 'Aucun front pendant bagotement');
ADVANCE_TIME(10000000); fb();
        IF fb.RawX < 5000 THEN oscillationSeen := TRUE; END_IF;
        ASSERT_FALSE(fb.RawButton, 'Aucun front pendant bagotement');
ADVANCE_TIME(10000000); fb();
        IF fb.RawX < 5000 THEN oscillationSeen := TRUE; END_IF;
        ASSERT_FALSE(fb.RawButton, 'Aucun front pendant bagotement');
ADVANCE_TIME(10000000); fb();
        IF fb.RawX < 5000 THEN oscillationSeen := TRUE; END_IF;
        ASSERT_FALSE(fb.RawButton, 'Aucun front pendant bagotement');
ADVANCE_TIME(10000000); fb();
        IF fb.RawX < 5000 THEN oscillationSeen := TRUE; END_IF;
        ASSERT_FALSE(fb.RawButton, 'Aucun front pendant bagotement');
ADVANCE_TIME(10000000); fb();
        IF fb.RawX < 5000 THEN oscillationSeen := TRUE; END_IF;
        ASSERT_FALSE(fb.RawButton, 'Aucun front pendant bagotement');
ADVANCE_TIME(10000000); fb();
        IF fb.RawX < 5000 THEN oscillationSeen := TRUE; END_IF;
        ASSERT_FALSE(fb.RawButton, 'Aucun front pendant bagotement');
ADVANCE_TIME(10000000); fb();
        IF fb.RawX < 5000 THEN oscillationSeen := TRUE; END_IF;
        ASSERT_FALSE(fb.RawButton, 'Aucun front pendant bagotement');
ADVANCE_TIME(10000000); fb();
        IF fb.RawX < 5000 THEN oscillationSeen := TRUE; END_IF;
        ASSERT_FALSE(fb.RawButton, 'Aucun front pendant bagotement');
ADVANCE_TIME(10000000); fb();
        IF fb.RawX < 5000 THEN oscillationSeen := TRUE; END_IF;
        ASSERT_FALSE(fb.RawButton, 'Aucun front pendant bagotement');
ADVANCE_TIME(10000000); fb();
        IF fb.RawX < 5000 THEN oscillationSeen := TRUE; END_IF;
        ASSERT_FALSE(fb.RawButton, 'Aucun front pendant bagotement');
ADVANCE_TIME(10000000); fb();
        IF fb.RawX < 5000 THEN oscillationSeen := TRUE; END_IF;
        ASSERT_FALSE(fb.RawButton, 'Aucun front pendant bagotement');
ADVANCE_TIME(10000000); fb();
        IF fb.RawX < 5000 THEN oscillationSeen := TRUE; END_IF;
        ASSERT_FALSE(fb.RawButton, 'Aucun front pendant bagotement');
ADVANCE_TIME(10000000); fb();
        IF fb.RawX < 5000 THEN oscillationSeen := TRUE; END_IF;
        ASSERT_FALSE(fb.RawButton, 'Aucun front pendant bagotement');
ADVANCE_TIME(10000000); fb();
        IF fb.RawX < 5000 THEN oscillationSeen := TRUE; END_IF;
        ASSERT_FALSE(fb.RawButton, 'Aucun front pendant bagotement');
ADVANCE_TIME(10000000); fb();
        IF fb.RawX < 5000 THEN oscillationSeen := TRUE; END_IF;
        ASSERT_FALSE(fb.RawButton, 'Aucun front pendant bagotement');
ADVANCE_TIME(10000000); fb();
        IF fb.RawX < 5000 THEN oscillationSeen := TRUE; END_IF;
        ASSERT_FALSE(fb.RawButton, 'Aucun front pendant bagotement');
ADVANCE_TIME(10000000); fb();
        IF fb.RawX < 5000 THEN oscillationSeen := TRUE; END_IF;
        ASSERT_FALSE(fb.RawButton, 'Aucun front pendant bagotement');
ADVANCE_TIME(10000000); fb();
        IF fb.RawX < 5000 THEN oscillationSeen := TRUE; END_IF;
        ASSERT_FALSE(fb.RawButton, 'Aucun front pendant bagotement');
ADVANCE_TIME(10000000); fb();
        IF fb.RawX < 5000 THEN oscillationSeen := TRUE; END_IF;
        ASSERT_FALSE(fb.RawButton, 'Aucun front pendant bagotement');
ADVANCE_TIME(10000000); fb();
        IF fb.RawX < 5000 THEN oscillationSeen := TRUE; END_IF;
        ASSERT_FALSE(fb.RawButton, 'Aucun front pendant bagotement');
ADVANCE_TIME(10000000); fb();
        IF fb.RawX < 5000 THEN oscillationSeen := TRUE; END_IF;
        ASSERT_FALSE(fb.RawButton, 'Aucun front pendant bagotement');
ADVANCE_TIME(10000000); fb();
        IF fb.RawX < 5000 THEN oscillationSeen := TRUE; END_IF;
        ASSERT_FALSE(fb.RawButton, 'Aucun front pendant bagotement');
ADVANCE_TIME(10000000); fb();
        IF fb.RawX < 5000 THEN oscillationSeen := TRUE; END_IF;
        ASSERT_FALSE(fb.RawButton, 'Aucun front pendant bagotement');
ADVANCE_TIME(10000000); fb();
        IF fb.RawX < 5000 THEN oscillationSeen := TRUE; END_IF;
        ASSERT_FALSE(fb.RawButton, 'Aucun front pendant bagotement');
ADVANCE_TIME(10000000); fb();
        IF fb.RawX < 5000 THEN oscillationSeen := TRUE; END_IF;
        ASSERT_FALSE(fb.RawButton, 'Aucun front pendant bagotement');
ADVANCE_TIME(10000000); fb();
        IF fb.RawX < 5000 THEN oscillationSeen := TRUE; END_IF;
        ASSERT_FALSE(fb.RawButton, 'Aucun front pendant bagotement');
ADVANCE_TIME(10000000); fb();
        IF fb.RawX < 5000 THEN oscillationSeen := TRUE; END_IF;
        ASSERT_FALSE(fb.RawButton, 'Aucun front pendant bagotement');
ADVANCE_TIME(10000000); fb();
        IF fb.RawX < 5000 THEN oscillationSeen := TRUE; END_IF;
        ASSERT_FALSE(fb.RawButton, 'Aucun front pendant bagotement');
ADVANCE_TIME(10000000); fb();
        IF fb.RawX < 5000 THEN oscillationSeen := TRUE; END_IF;
        ASSERT_FALSE(fb.RawButton, 'Aucun front pendant bagotement');
ADVANCE_TIME(10000000); fb();
        IF fb.RawX < 5000 THEN oscillationSeen := TRUE; END_IF;
        ASSERT_FALSE(fb.RawButton, 'Aucun front pendant bagotement');
ADVANCE_TIME(10000000); fb();
        IF fb.RawX < 5000 THEN oscillationSeen := TRUE; END_IF;
        ASSERT_FALSE(fb.RawButton, 'Aucun front pendant bagotement');
ADVANCE_TIME(10000000); fb();
        IF fb.RawX < 5000 THEN oscillationSeen := TRUE; END_IF;
        ASSERT_FALSE(fb.RawButton, 'Aucun front pendant bagotement');
ADVANCE_TIME(10000000); fb();
        IF fb.RawX < 5000 THEN oscillationSeen := TRUE; END_IF;
        ASSERT_FALSE(fb.RawButton, 'Aucun front pendant bagotement');
ADVANCE_TIME(10000000); fb();
        IF fb.RawX < 5000 THEN oscillationSeen := TRUE; END_IF;
        ASSERT_FALSE(fb.RawButton, 'Aucun front pendant bagotement');
ADVANCE_TIME(10000000); fb();
        IF fb.RawX < 5000 THEN oscillationSeen := TRUE; END_IF;
        ASSERT_FALSE(fb.RawButton, 'Aucun front pendant bagotement');
ADVANCE_TIME(10000000); fb();
        IF fb.RawX < 5000 THEN oscillationSeen := TRUE; END_IF;
        ASSERT_FALSE(fb.RawButton, 'Aucun front pendant bagotement');
ADVANCE_TIME(10000000); fb();
        IF fb.RawX < 5000 THEN oscillationSeen := TRUE; END_IF;
        ASSERT_FALSE(fb.RawButton, 'Aucun front pendant bagotement');
ADVANCE_TIME(10000000); fb();
        IF fb.RawX < 5000 THEN oscillationSeen := TRUE; END_IF;
        ASSERT_FALSE(fb.RawButton, 'Aucun front pendant bagotement');
ADVANCE_TIME(10000000); fb();
        IF fb.RawX < 5000 THEN oscillationSeen := TRUE; END_IF;
        ASSERT_FALSE(fb.RawButton, 'Aucun front pendant bagotement');
ADVANCE_TIME(10000000); fb();
        IF fb.RawX < 5000 THEN oscillationSeen := TRUE; END_IF;
        ASSERT_FALSE(fb.RawButton, 'Aucun front pendant bagotement');
ADVANCE_TIME(10000000); fb();
        IF fb.RawX < 5000 THEN oscillationSeen := TRUE; END_IF;
        ASSERT_FALSE(fb.RawButton, 'Aucun front pendant bagotement');
ADVANCE_TIME(10000000); fb();
        IF fb.RawX < 5000 THEN oscillationSeen := TRUE; END_IF;
        ASSERT_FALSE(fb.RawButton, 'Aucun front pendant bagotement');
ADVANCE_TIME(10000000); fb();
        IF fb.RawX < 5000 THEN oscillationSeen := TRUE; END_IF;
        ASSERT_FALSE(fb.RawButton, 'Aucun front pendant bagotement');
ADVANCE_TIME(10000000); fb();
        IF fb.RawX < 5000 THEN oscillationSeen := TRUE; END_IF;
        ASSERT_FALSE(fb.RawButton, 'Aucun front pendant bagotement');
ADVANCE_TIME(10000000); fb();
        IF fb.RawX < 5000 THEN oscillationSeen := TRUE; END_IF;
        ASSERT_FALSE(fb.RawButton, 'Aucun front pendant bagotement');
ADVANCE_TIME(10000000); fb();
        IF fb.RawX < 5000 THEN oscillationSeen := TRUE; END_IF;
        ASSERT_FALSE(fb.RawButton, 'Aucun front pendant bagotement');
ADVANCE_TIME(10000000); fb();
        IF fb.RawX < 5000 THEN oscillationSeen := TRUE; END_IF;
        ASSERT_FALSE(fb.RawButton, 'Aucun front pendant bagotement');
ADVANCE_TIME(10000000); fb();
        IF fb.RawX < 5000 THEN oscillationSeen := TRUE; END_IF;
        ASSERT_FALSE(fb.RawButton, 'Aucun front pendant bagotement');
ADVANCE_TIME(10000000); fb();
        IF fb.RawX < 5000 THEN oscillationSeen := TRUE; END_IF;
        ASSERT_FALSE(fb.RawButton, 'Aucun front pendant bagotement');
ADVANCE_TIME(10000000); fb();
        IF fb.RawX < 5000 THEN oscillationSeen := TRUE; END_IF;
        ASSERT_FALSE(fb.RawButton, 'Aucun front pendant bagotement');
ADVANCE_TIME(10000000); fb();
        IF fb.RawX < 5000 THEN oscillationSeen := TRUE; END_IF;
        ASSERT_FALSE(fb.RawButton, 'Aucun front pendant bagotement');
ADVANCE_TIME(10000000); fb();
        IF fb.RawX < 5000 THEN oscillationSeen := TRUE; END_IF;
        ASSERT_FALSE(fb.RawButton, 'Aucun front pendant bagotement');
ADVANCE_TIME(10000000); fb();
        IF fb.RawX < 5000 THEN oscillationSeen := TRUE; END_IF;
        ASSERT_FALSE(fb.RawButton, 'Aucun front pendant bagotement');
ADVANCE_TIME(10000000); fb();
        IF fb.RawX < 5000 THEN oscillationSeen := TRUE; END_IF;
        ASSERT_FALSE(fb.RawButton, 'Aucun front pendant bagotement');
ADVANCE_TIME(10000000); fb();
        IF fb.RawX < 5000 THEN oscillationSeen := TRUE; END_IF;
        ASSERT_FALSE(fb.RawButton, 'Aucun front pendant bagotement');
ADVANCE_TIME(10000000); fb();
        IF fb.RawX < 5000 THEN oscillationSeen := TRUE; END_IF;
        ASSERT_FALSE(fb.RawButton, 'Aucun front pendant bagotement');
ADVANCE_TIME(10000000); fb();
        IF fb.RawX < 5000 THEN oscillationSeen := TRUE; END_IF;
        ASSERT_FALSE(fb.RawButton, 'Aucun front pendant bagotement');
ADVANCE_TIME(10000000); fb();
        IF fb.RawX < 5000 THEN oscillationSeen := TRUE; END_IF;
        ASSERT_FALSE(fb.RawButton, 'Aucun front pendant bagotement');
ADVANCE_TIME(10000000); fb();
        IF fb.RawX < 5000 THEN oscillationSeen := TRUE; END_IF;
        ASSERT_FALSE(fb.RawButton, 'Aucun front pendant bagotement');
ADVANCE_TIME(10000000); fb();
        IF fb.RawX < 5000 THEN oscillationSeen := TRUE; END_IF;
        ASSERT_FALSE(fb.RawButton, 'Aucun front pendant bagotement');
ADVANCE_TIME(10000000); fb();
        IF fb.RawX < 5000 THEN oscillationSeen := TRUE; END_IF;
        ASSERT_FALSE(fb.RawButton, 'Aucun front pendant bagotement');
ADVANCE_TIME(10000000); fb();
        IF fb.RawX < 5000 THEN oscillationSeen := TRUE; END_IF;
        ASSERT_FALSE(fb.RawButton, 'Aucun front pendant bagotement');
ADVANCE_TIME(10000000); fb();
        IF fb.RawX < 5000 THEN oscillationSeen := TRUE; END_IF;
        ASSERT_FALSE(fb.RawButton, 'Aucun front pendant bagotement');
ADVANCE_TIME(10000000); fb();
        IF fb.RawX < 5000 THEN oscillationSeen := TRUE; END_IF;
        ASSERT_FALSE(fb.RawButton, 'Aucun front pendant bagotement');
ADVANCE_TIME(10000000); fb();
        IF fb.RawX < 5000 THEN oscillationSeen := TRUE; END_IF;
        ASSERT_FALSE(fb.RawButton, 'Aucun front pendant bagotement');
ADVANCE_TIME(10000000); fb();
        IF fb.RawX < 5000 THEN oscillationSeen := TRUE; END_IF;
        ASSERT_FALSE(fb.RawButton, 'Aucun front pendant bagotement');
ADVANCE_TIME(10000000); fb();
        IF fb.RawX < 5000 THEN oscillationSeen := TRUE; END_IF;
        ASSERT_FALSE(fb.RawButton, 'Aucun front pendant bagotement');
ADVANCE_TIME(10000000); fb();
        IF fb.RawX < 5000 THEN oscillationSeen := TRUE; END_IF;
        ASSERT_FALSE(fb.RawButton, 'Aucun front pendant bagotement');
ADVANCE_TIME(10000000); fb();
        IF fb.RawX < 5000 THEN oscillationSeen := TRUE; END_IF;
        ASSERT_FALSE(fb.RawButton, 'Aucun front pendant bagotement');
ADVANCE_TIME(10000000); fb();
        IF fb.RawX < 5000 THEN oscillationSeen := TRUE; END_IF;
        ASSERT_FALSE(fb.RawButton, 'Aucun front pendant bagotement');
ADVANCE_TIME(10000000); fb();
        IF fb.RawX < 5000 THEN oscillationSeen := TRUE; END_IF;
        ASSERT_FALSE(fb.RawButton, 'Aucun front pendant bagotement');
ADVANCE_TIME(10000000); fb();
        IF fb.RawX < 5000 THEN oscillationSeen := TRUE; END_IF;
        ASSERT_FALSE(fb.RawButton, 'Aucun front pendant bagotement');
ADVANCE_TIME(10000000); fb();
        IF fb.RawX < 5000 THEN oscillationSeen := TRUE; END_IF;
        ASSERT_FALSE(fb.RawButton, 'Aucun front pendant bagotement');
ADVANCE_TIME(10000000); fb();
        IF fb.RawX < 5000 THEN oscillationSeen := TRUE; END_IF;
        ASSERT_FALSE(fb.RawButton, 'Aucun front pendant bagotement');
ADVANCE_TIME(10000000); fb();
        IF fb.RawX < 5000 THEN oscillationSeen := TRUE; END_IF;
        ASSERT_FALSE(fb.RawButton, 'Aucun front pendant bagotement');
ADVANCE_TIME(10000000); fb();
        IF fb.RawX < 5000 THEN oscillationSeen := TRUE; END_IF;
        ASSERT_FALSE(fb.RawButton, 'Aucun front pendant bagotement');
ADVANCE_TIME(10000000); fb();
        IF fb.RawX < 5000 THEN oscillationSeen := TRUE; END_IF;
        ASSERT_FALSE(fb.RawButton, 'Aucun front pendant bagotement');
ADVANCE_TIME(10000000); fb();
        IF fb.RawX < 5000 THEN oscillationSeen := TRUE; END_IF;
        ASSERT_FALSE(fb.RawButton, 'Aucun front pendant bagotement');
ADVANCE_TIME(10000000); fb();
        IF fb.RawX < 5000 THEN oscillationSeen := TRUE; END_IF;
        ASSERT_FALSE(fb.RawButton, 'Aucun front pendant bagotement');
ADVANCE_TIME(10000000); fb();
        IF fb.RawX < 5000 THEN oscillationSeen := TRUE; END_IF;
        ASSERT_FALSE(fb.RawButton, 'Aucun front pendant bagotement');
ADVANCE_TIME(10000000); fb();
        IF fb.RawX < 5000 THEN oscillationSeen := TRUE; END_IF;
        ASSERT_FALSE(fb.RawButton, 'Aucun front pendant bagotement');
ADVANCE_TIME(10000000); fb();
        IF fb.RawX < 5000 THEN oscillationSeen := TRUE; END_IF;
        ASSERT_FALSE(fb.RawButton, 'Aucun front pendant bagotement');
ADVANCE_TIME(10000000); fb();
        IF fb.RawX < 5000 THEN oscillationSeen := TRUE; END_IF;
        ASSERT_FALSE(fb.RawButton, 'Aucun front pendant bagotement');
ADVANCE_TIME(10000000); fb();
        IF fb.RawX < 5000 THEN oscillationSeen := TRUE; END_IF;
        ASSERT_FALSE(fb.RawButton, 'Aucun front pendant bagotement');
ADVANCE_TIME(10000000); fb();
        IF fb.RawX < 5000 THEN oscillationSeen := TRUE; END_IF;
        ASSERT_FALSE(fb.RawButton, 'Aucun front pendant bagotement');
ADVANCE_TIME(10000000); fb();
        IF fb.RawX < 5000 THEN oscillationSeen := TRUE; END_IF;
        ASSERT_FALSE(fb.RawButton, 'Aucun front pendant bagotement');
ADVANCE_TIME(10000000); fb();
        IF fb.RawX < 5000 THEN oscillationSeen := TRUE; END_IF;
        ASSERT_FALSE(fb.RawButton, 'Aucun front pendant bagotement');
ADVANCE_TIME(10000000); fb();
        IF fb.RawX < 5000 THEN oscillationSeen := TRUE; END_IF;
        ASSERT_FALSE(fb.RawButton, 'Aucun front pendant bagotement');
ADVANCE_TIME(10000000); fb();
        IF fb.RawX < 5000 THEN oscillationSeen := TRUE; END_IF;
        ASSERT_FALSE(fb.RawButton, 'Aucun front pendant bagotement');
ADVANCE_TIME(10000000); fb();
        IF fb.RawX < 5000 THEN oscillationSeen := TRUE; END_IF;
        ASSERT_FALSE(fb.RawButton, 'Aucun front pendant bagotement');
ADVANCE_TIME(10000000); fb();
        IF fb.RawX < 5000 THEN oscillationSeen := TRUE; END_IF;
        ASSERT_FALSE(fb.RawButton, 'Aucun front pendant bagotement');
ADVANCE_TIME(10000000); fb();
        IF fb.RawX < 5000 THEN oscillationSeen := TRUE; END_IF;
        ASSERT_FALSE(fb.RawButton, 'Aucun front pendant bagotement');
ADVANCE_TIME(10000000); fb();
        IF fb.RawX < 5000 THEN oscillationSeen := TRUE; END_IF;
        ASSERT_FALSE(fb.RawButton, 'Aucun front pendant bagotement');
ADVANCE_TIME(10000000); fb();
        IF fb.RawX < 5000 THEN oscillationSeen := TRUE; END_IF;
        ASSERT_FALSE(fb.RawButton, 'Aucun front pendant bagotement');
ADVANCE_TIME(10000000); fb();
        IF fb.RawX < 5000 THEN oscillationSeen := TRUE; END_IF;
        ASSERT_FALSE(fb.RawButton, 'Aucun front pendant bagotement');
ADVANCE_TIME(10000000); fb();
        IF fb.RawX < 5000 THEN oscillationSeen := TRUE; END_IF;
        ASSERT_FALSE(fb.RawButton, 'Aucun front pendant bagotement');
ADVANCE_TIME(10000000); fb();
        IF fb.RawX < 5000 THEN oscillationSeen := TRUE; END_IF;
        ASSERT_FALSE(fb.RawButton, 'Aucun front pendant bagotement');
ADVANCE_TIME(10000000); fb();
        IF fb.RawX < 5000 THEN oscillationSeen := TRUE; END_IF;
        ASSERT_FALSE(fb.RawButton, 'Aucun front pendant bagotement');
ADVANCE_TIME(10000000); fb();
        IF fb.RawX < 5000 THEN oscillationSeen := TRUE; END_IF;
        ASSERT_FALSE(fb.RawButton, 'Aucun front pendant bagotement');
ADVANCE_TIME(10000000); fb();
        IF fb.RawX < 5000 THEN oscillationSeen := TRUE; END_IF;
        ASSERT_FALSE(fb.RawButton, 'Aucun front pendant bagotement');
ADVANCE_TIME(10000000); fb();
        IF fb.RawX < 5000 THEN oscillationSeen := TRUE; END_IF;
        ASSERT_FALSE(fb.RawButton, 'Aucun front pendant bagotement');
ADVANCE_TIME(10000000); fb();
        IF fb.RawX < 5000 THEN oscillationSeen := TRUE; END_IF;
        ASSERT_FALSE(fb.RawButton, 'Aucun front pendant bagotement');
ADVANCE_TIME(10000000); fb();
        IF fb.RawX < 5000 THEN oscillationSeen := TRUE; END_IF;
        ASSERT_FALSE(fb.RawButton, 'Aucun front pendant bagotement');
ADVANCE_TIME(10000000); fb();
        IF fb.RawX < 5000 THEN oscillationSeen := TRUE; END_IF;
        ASSERT_FALSE(fb.RawButton, 'Aucun front pendant bagotement');
ADVANCE_TIME(10000000); fb();
        IF fb.RawX < 5000 THEN oscillationSeen := TRUE; END_IF;
        ASSERT_FALSE(fb.RawButton, 'Aucun front pendant bagotement');
ADVANCE_TIME(10000000); fb();
        IF fb.RawX < 5000 THEN oscillationSeen := TRUE; END_IF;
        ASSERT_FALSE(fb.RawButton, 'Aucun front pendant bagotement');
ADVANCE_TIME(10000000); fb();
        IF fb.RawX < 5000 THEN oscillationSeen := TRUE; END_IF;
        ASSERT_FALSE(fb.RawButton, 'Aucun front pendant bagotement');
ADVANCE_TIME(10000000); fb();
        IF fb.RawX < 5000 THEN oscillationSeen := TRUE; END_IF;
        ASSERT_FALSE(fb.RawButton, 'Aucun front pendant bagotement');
ADVANCE_TIME(10000000); fb();
        IF fb.RawX < 5000 THEN oscillationSeen := TRUE; END_IF;
        ASSERT_FALSE(fb.RawButton, 'Aucun front pendant bagotement');
ADVANCE_TIME(10000000); fb();
        IF fb.RawX < 5000 THEN oscillationSeen := TRUE; END_IF;
        ASSERT_FALSE(fb.RawButton, 'Aucun front pendant bagotement');
ADVANCE_TIME(10000000); fb();
        IF fb.RawX < 5000 THEN oscillationSeen := TRUE; END_IF;
        ASSERT_FALSE(fb.RawButton, 'Aucun front pendant bagotement');
ADVANCE_TIME(10000000); fb();
        IF fb.RawX < 5000 THEN oscillationSeen := TRUE; END_IF;
        ASSERT_FALSE(fb.RawButton, 'Aucun front pendant bagotement');
ADVANCE_TIME(10000000); fb();
        IF fb.RawX < 5000 THEN oscillationSeen := TRUE; END_IF;
        ASSERT_FALSE(fb.RawButton, 'Aucun front pendant bagotement');
ADVANCE_TIME(10000000); fb();
        IF fb.RawX < 5000 THEN oscillationSeen := TRUE; END_IF;
        ASSERT_FALSE(fb.RawButton, 'Aucun front pendant bagotement');
ADVANCE_TIME(10000000); fb();
        IF fb.RawX < 5000 THEN oscillationSeen := TRUE; END_IF;
        ASSERT_FALSE(fb.RawButton, 'Aucun front pendant bagotement');
ADVANCE_TIME(10000000); fb();
        IF fb.RawX < 5000 THEN oscillationSeen := TRUE; END_IF;
        ASSERT_FALSE(fb.RawButton, 'Aucun front pendant bagotement');
ADVANCE_TIME(10000000); fb();
        IF fb.RawX < 5000 THEN oscillationSeen := TRUE; END_IF;
        ASSERT_FALSE(fb.RawButton, 'Aucun front pendant bagotement');
ADVANCE_TIME(10000000); fb();
        IF fb.RawX < 5000 THEN oscillationSeen := TRUE; END_IF;
        ASSERT_FALSE(fb.RawButton, 'Aucun front pendant bagotement');
ADVANCE_TIME(10000000); fb();
        IF fb.RawX < 5000 THEN oscillationSeen := TRUE; END_IF;
        ASSERT_FALSE(fb.RawButton, 'Aucun front pendant bagotement');
ADVANCE_TIME(10000000); fb();
        IF fb.RawX < 5000 THEN oscillationSeen := TRUE; END_IF;
        ASSERT_FALSE(fb.RawButton, 'Aucun front pendant bagotement');
ADVANCE_TIME(10000000); fb();
        IF fb.RawX < 5000 THEN oscillationSeen := TRUE; END_IF;
        ASSERT_FALSE(fb.RawButton, 'Aucun front pendant bagotement');
ADVANCE_TIME(10000000); fb();
        IF fb.RawX < 5000 THEN oscillationSeen := TRUE; END_IF;
        ASSERT_FALSE(fb.RawButton, 'Aucun front pendant bagotement');
ADVANCE_TIME(10000000); fb();
        IF fb.RawX < 5000 THEN oscillationSeen := TRUE; END_IF;
        ASSERT_FALSE(fb.RawButton, 'Aucun front pendant bagotement');
ADVANCE_TIME(10000000); fb();
        IF fb.RawX < 5000 THEN oscillationSeen := TRUE; END_IF;
        ASSERT_FALSE(fb.RawButton, 'Aucun front pendant bagotement');
ADVANCE_TIME(10000000); fb();
        IF fb.RawX < 5000 THEN oscillationSeen := TRUE; END_IF;
        ASSERT_FALSE(fb.RawButton, 'Aucun front pendant bagotement');
ADVANCE_TIME(10000000); fb();
        IF fb.RawX < 5000 THEN oscillationSeen := TRUE; END_IF;
        ASSERT_FALSE(fb.RawButton, 'Aucun front pendant bagotement');
ADVANCE_TIME(10000000); fb();
        IF fb.RawX < 5000 THEN oscillationSeen := TRUE; END_IF;
        ASSERT_FALSE(fb.RawButton, 'Aucun front pendant bagotement');
ADVANCE_TIME(10000000); fb();
        IF fb.RawX < 5000 THEN oscillationSeen := TRUE; END_IF;
        ASSERT_FALSE(fb.RawButton, 'Aucun front pendant bagotement');
ADVANCE_TIME(10000000); fb();
        IF fb.RawX < 5000 THEN oscillationSeen := TRUE; END_IF;
        ASSERT_FALSE(fb.RawButton, 'Aucun front pendant bagotement');
ADVANCE_TIME(10000000); fb();
        IF fb.RawX < 5000 THEN oscillationSeen := TRUE; END_IF;
        ASSERT_FALSE(fb.RawButton, 'Aucun front pendant bagotement');
ADVANCE_TIME(10000000); fb();
        IF fb.RawX < 5000 THEN oscillationSeen := TRUE; END_IF;
        ASSERT_FALSE(fb.RawButton, 'Aucun front pendant bagotement');
ADVANCE_TIME(10000000); fb();
        IF fb.RawX < 5000 THEN oscillationSeen := TRUE; END_IF;
        ASSERT_FALSE(fb.RawButton, 'Aucun front pendant bagotement');
ADVANCE_TIME(10000000); fb();
        IF fb.RawX < 5000 THEN oscillationSeen := TRUE; END_IF;
        ASSERT_FALSE(fb.RawButton, 'Aucun front pendant bagotement');
ADVANCE_TIME(10000000); fb();
        IF fb.RawX < 5000 THEN oscillationSeen := TRUE; END_IF;
        ASSERT_FALSE(fb.RawButton, 'Aucun front pendant bagotement');
ADVANCE_TIME(10000000); fb();
        IF fb.RawX < 5000 THEN oscillationSeen := TRUE; END_IF;
        ASSERT_FALSE(fb.RawButton, 'Aucun front pendant bagotement');
ADVANCE_TIME(10000000); fb();
        IF fb.RawX < 5000 THEN oscillationSeen := TRUE; END_IF;
        ASSERT_FALSE(fb.RawButton, 'Aucun front pendant bagotement');
ADVANCE_TIME(10000000); fb();
        IF fb.RawX < 5000 THEN oscillationSeen := TRUE; END_IF;
        ASSERT_FALSE(fb.RawButton, 'Aucun front pendant bagotement');
ADVANCE_TIME(10000000); fb();
        IF fb.RawX < 5000 THEN oscillationSeen := TRUE; END_IF;
        ASSERT_FALSE(fb.RawButton, 'Aucun front pendant bagotement');
ADVANCE_TIME(10000000); fb();
        IF fb.RawX < 5000 THEN oscillationSeen := TRUE; END_IF;
        ASSERT_FALSE(fb.RawButton, 'Aucun front pendant bagotement');
ADVANCE_TIME(10000000); fb();
        IF fb.RawX < 5000 THEN oscillationSeen := TRUE; END_IF;
        ASSERT_FALSE(fb.RawButton, 'Aucun front pendant bagotement');
ADVANCE_TIME(10000000); fb();
        IF fb.RawX < 5000 THEN oscillationSeen := TRUE; END_IF;
        ASSERT_FALSE(fb.RawButton, 'Aucun front pendant bagotement');
ADVANCE_TIME(10000000); fb();
        IF fb.RawX < 5000 THEN oscillationSeen := TRUE; END_IF;
        ASSERT_FALSE(fb.RawButton, 'Aucun front pendant bagotement');
ADVANCE_TIME(10000000); fb();
        IF fb.RawX < 5000 THEN oscillationSeen := TRUE; END_IF;
        ASSERT_FALSE(fb.RawButton, 'Aucun front pendant bagotement');
ADVANCE_TIME(10000000); fb();
        IF fb.RawX < 5000 THEN oscillationSeen := TRUE; END_IF;
        ASSERT_FALSE(fb.RawButton, 'Aucun front pendant bagotement');
ADVANCE_TIME(10000000); fb();
        IF fb.RawX < 5000 THEN oscillationSeen := TRUE; END_IF;
        ASSERT_FALSE(fb.RawButton, 'Aucun front pendant bagotement');
ADVANCE_TIME(10000000); fb();
        IF fb.RawX < 5000 THEN oscillationSeen := TRUE; END_IF;
        ASSERT_FALSE(fb.RawButton, 'Aucun front pendant bagotement');
ADVANCE_TIME(10000000); fb();
        IF fb.RawX < 5000 THEN oscillationSeen := TRUE; END_IF;
        ASSERT_FALSE(fb.RawButton, 'Aucun front pendant bagotement');
ADVANCE_TIME(10000000); fb();
        IF fb.RawX < 5000 THEN oscillationSeen := TRUE; END_IF;
        ASSERT_FALSE(fb.RawButton, 'Aucun front pendant bagotement');
ADVANCE_TIME(10000000); fb();
        IF fb.RawX < 5000 THEN oscillationSeen := TRUE; END_IF;
        ASSERT_FALSE(fb.RawButton, 'Aucun front pendant bagotement');
ADVANCE_TIME(10000000); fb();
        IF fb.RawX < 5000 THEN oscillationSeen := TRUE; END_IF;
        ASSERT_FALSE(fb.RawButton, 'Aucun front pendant bagotement');
ADVANCE_TIME(10000000); fb();
        IF fb.RawX < 5000 THEN oscillationSeen := TRUE; END_IF;
        ASSERT_FALSE(fb.RawButton, 'Aucun front pendant bagotement');
ADVANCE_TIME(10000000); fb();
        IF fb.RawX < 5000 THEN oscillationSeen := TRUE; END_IF;
        ASSERT_FALSE(fb.RawButton, 'Aucun front pendant bagotement');
ADVANCE_TIME(10000000); fb();
        IF fb.RawX < 5000 THEN oscillationSeen := TRUE; END_IF;
        ASSERT_FALSE(fb.RawButton, 'Aucun front pendant bagotement');
ADVANCE_TIME(10000000); fb();
        IF fb.RawX < 5000 THEN oscillationSeen := TRUE; END_IF;
        ASSERT_FALSE(fb.RawButton, 'Aucun front pendant bagotement');
ADVANCE_TIME(10000000); fb();
        IF fb.RawX < 5000 THEN oscillationSeen := TRUE; END_IF;
        ASSERT_FALSE(fb.RawButton, 'Aucun front pendant bagotement');
ADVANCE_TIME(10000000); fb();
        IF fb.RawX < 5000 THEN oscillationSeen := TRUE; END_IF;
        ASSERT_FALSE(fb.RawButton, 'Aucun front pendant bagotement');
ADVANCE_TIME(10000000); fb();
        IF fb.RawX < 5000 THEN oscillationSeen := TRUE; END_IF;
        ASSERT_FALSE(fb.RawButton, 'Aucun front pendant bagotement');
ADVANCE_TIME(10000000); fb();
        IF fb.RawX < 5000 THEN oscillationSeen := TRUE; END_IF;
        ASSERT_FALSE(fb.RawButton, 'Aucun front pendant bagotement');
ADVANCE_TIME(10000000); fb();
        IF fb.RawX < 5000 THEN oscillationSeen := TRUE; END_IF;
        ASSERT_FALSE(fb.RawButton, 'Aucun front pendant bagotement');
ADVANCE_TIME(10000000); fb();
        IF fb.RawX < 5000 THEN oscillationSeen := TRUE; END_IF;
        ASSERT_FALSE(fb.RawButton, 'Aucun front pendant bagotement');
ADVANCE_TIME(10000000); fb();
        IF fb.RawX < 5000 THEN oscillationSeen := TRUE; END_IF;
        ASSERT_FALSE(fb.RawButton, 'Aucun front pendant bagotement');
ADVANCE_TIME(10000000); fb();
        IF fb.RawX < 5000 THEN oscillationSeen := TRUE; END_IF;
        ASSERT_FALSE(fb.RawButton, 'Aucun front pendant bagotement');
ADVANCE_TIME(10000000); fb();
        IF fb.RawX < 5000 THEN oscillationSeen := TRUE; END_IF;
        ASSERT_FALSE(fb.RawButton, 'Aucun front pendant bagotement');
ADVANCE_TIME(10000000); fb();
        IF fb.RawX < 5000 THEN oscillationSeen := TRUE; END_IF;
        ASSERT_FALSE(fb.RawButton, 'Aucun front pendant bagotement');
ADVANCE_TIME(10000000); fb();
        IF fb.RawX < 5000 THEN oscillationSeen := TRUE; END_IF;
        ASSERT_FALSE(fb.RawButton, 'Aucun front pendant bagotement');
ADVANCE_TIME(10000000); fb();
        IF fb.RawX < 5000 THEN oscillationSeen := TRUE; END_IF;
        ASSERT_FALSE(fb.RawButton, 'Aucun front pendant bagotement');
ADVANCE_TIME(10000000); fb();
        IF fb.RawX < 5000 THEN oscillationSeen := TRUE; END_IF;
        ASSERT_FALSE(fb.RawButton, 'Aucun front pendant bagotement');
ADVANCE_TIME(10000000); fb();
        IF fb.RawX < 5000 THEN oscillationSeen := TRUE; END_IF;
        ASSERT_FALSE(fb.RawButton, 'Aucun front pendant bagotement');
ADVANCE_TIME(10000000); fb();
        IF fb.RawX < 5000 THEN oscillationSeen := TRUE; END_IF;
        ASSERT_FALSE(fb.RawButton, 'Aucun front pendant bagotement');
ADVANCE_TIME(10000000); fb();
        IF fb.RawX < 5000 THEN oscillationSeen := TRUE; END_IF;
        ASSERT_FALSE(fb.RawButton, 'Aucun front pendant bagotement');
ADVANCE_TIME(10000000); fb();
        IF fb.RawX < 5000 THEN oscillationSeen := TRUE; END_IF;
        ASSERT_FALSE(fb.RawButton, 'Aucun front pendant bagotement');
ADVANCE_TIME(10000000); fb();
        IF fb.RawX < 5000 THEN oscillationSeen := TRUE; END_IF;
        ASSERT_FALSE(fb.RawButton, 'Aucun front pendant bagotement');
ADVANCE_TIME(10000000); fb();
        IF fb.RawX < 5000 THEN oscillationSeen := TRUE; END_IF;
        ASSERT_FALSE(fb.RawButton, 'Aucun front pendant bagotement');
ADVANCE_TIME(10000000); fb();
        IF fb.RawX < 5000 THEN oscillationSeen := TRUE; END_IF;
        ASSERT_FALSE(fb.RawButton, 'Aucun front pendant bagotement');
ADVANCE_TIME(10000000); fb();
        IF fb.RawX < 5000 THEN oscillationSeen := TRUE; END_IF;
        ASSERT_FALSE(fb.RawButton, 'Aucun front pendant bagotement');
ADVANCE_TIME(10000000); fb();
        IF fb.RawX < 5000 THEN oscillationSeen := TRUE; END_IF;
        ASSERT_FALSE(fb.RawButton, 'Aucun front pendant bagotement');
ADVANCE_TIME(10000000); fb();
        IF fb.RawX < 5000 THEN oscillationSeen := TRUE; END_IF;
        ASSERT_FALSE(fb.RawButton, 'Aucun front pendant bagotement');
ADVANCE_TIME(10000000); fb();
        IF fb.RawX < 5000 THEN oscillationSeen := TRUE; END_IF;
        ASSERT_FALSE(fb.RawButton, 'Aucun front pendant bagotement');
ADVANCE_TIME(10000000); fb();
        IF fb.RawX < 5000 THEN oscillationSeen := TRUE; END_IF;
        ASSERT_FALSE(fb.RawButton, 'Aucun front pendant bagotement');
ADVANCE_TIME(10000000); fb();
        IF fb.RawX < 5000 THEN oscillationSeen := TRUE; END_IF;
        ASSERT_FALSE(fb.RawButton, 'Aucun front pendant bagotement');
ADVANCE_TIME(10000000); fb();
        IF fb.RawX < 5000 THEN oscillationSeen := TRUE; END_IF;
        ASSERT_FALSE(fb.RawButton, 'Aucun front pendant bagotement');
ADVANCE_TIME(10000000); fb();
        IF fb.RawX < 5000 THEN oscillationSeen := TRUE; END_IF;
        ASSERT_FALSE(fb.RawButton, 'Aucun front pendant bagotement');
ADVANCE_TIME(10000000); fb();
        IF fb.RawX < 5000 THEN oscillationSeen := TRUE; END_IF;
        ASSERT_FALSE(fb.RawButton, 'Aucun front pendant bagotement');
ADVANCE_TIME(10000000); fb();
        IF fb.RawX < 5000 THEN oscillationSeen := TRUE; END_IF;
        ASSERT_FALSE(fb.RawButton, 'Aucun front pendant bagotement');
ADVANCE_TIME(10000000); fb();
        IF fb.RawX < 5000 THEN oscillationSeen := TRUE; END_IF;
        ASSERT_FALSE(fb.RawButton, 'Aucun front pendant bagotement');
ADVANCE_TIME(10000000); fb();
        IF fb.RawX < 5000 THEN oscillationSeen := TRUE; END_IF;
        ASSERT_FALSE(fb.RawButton, 'Aucun front pendant bagotement');
ADVANCE_TIME(10000000); fb();
        IF fb.RawX < 5000 THEN oscillationSeen := TRUE; END_IF;
        ASSERT_FALSE(fb.RawButton, 'Aucun front pendant bagotement');
ADVANCE_TIME(10000000); fb();
        IF fb.RawX < 5000 THEN oscillationSeen := TRUE; END_IF;
        ASSERT_FALSE(fb.RawButton, 'Aucun front pendant bagotement');
ADVANCE_TIME(10000000); fb();
        IF fb.RawX < 5000 THEN oscillationSeen := TRUE; END_IF;
        ASSERT_FALSE(fb.RawButton, 'Aucun front pendant bagotement');
ADVANCE_TIME(10000000); fb();
        IF fb.RawX < 5000 THEN oscillationSeen := TRUE; END_IF;
        ASSERT_FALSE(fb.RawButton, 'Aucun front pendant bagotement');
ADVANCE_TIME(10000000); fb();
        IF fb.RawX < 5000 THEN oscillationSeen := TRUE; END_IF;
        ASSERT_FALSE(fb.RawButton, 'Aucun front pendant bagotement');
ADVANCE_TIME(10000000); fb();
        IF fb.RawX < 5000 THEN oscillationSeen := TRUE; END_IF;
        ASSERT_FALSE(fb.RawButton, 'Aucun front pendant bagotement');
ADVANCE_TIME(10000000); fb();
        IF fb.RawX < 5000 THEN oscillationSeen := TRUE; END_IF;
        ASSERT_FALSE(fb.RawButton, 'Aucun front pendant bagotement');
ADVANCE_TIME(10000000); fb();
        IF fb.RawX < 5000 THEN oscillationSeen := TRUE; END_IF;
        ASSERT_FALSE(fb.RawButton, 'Aucun front pendant bagotement');
ADVANCE_TIME(10000000); fb();
        IF fb.RawX < 5000 THEN oscillationSeen := TRUE; END_IF;
        ASSERT_FALSE(fb.RawButton, 'Aucun front pendant bagotement');
ADVANCE_TIME(10000000); fb();
        IF fb.RawX < 5000 THEN oscillationSeen := TRUE; END_IF;
        ASSERT_FALSE(fb.RawButton, 'Aucun front pendant bagotement');
ADVANCE_TIME(10000000); fb();
        IF fb.RawX < 5000 THEN oscillationSeen := TRUE; END_IF;
        ASSERT_FALSE(fb.RawButton, 'Aucun front pendant bagotement');
ADVANCE_TIME(10000000); fb();
        IF fb.RawX < 5000 THEN oscillationSeen := TRUE; END_IF;
        ASSERT_FALSE(fb.RawButton, 'Aucun front pendant bagotement');
ADVANCE_TIME(10000000); fb();
        IF fb.RawX < 5000 THEN oscillationSeen := TRUE; END_IF;
        ASSERT_FALSE(fb.RawButton, 'Aucun front pendant bagotement');
ADVANCE_TIME(10000000); fb();
        IF fb.RawX < 5000 THEN oscillationSeen := TRUE; END_IF;
        ASSERT_FALSE(fb.RawButton, 'Aucun front pendant bagotement');
ADVANCE_TIME(10000000); fb();
        IF fb.RawX < 5000 THEN oscillationSeen := TRUE; END_IF;
        ASSERT_FALSE(fb.RawButton, 'Aucun front pendant bagotement');
ADVANCE_TIME(10000000); fb();
        IF fb.RawX < 5000 THEN oscillationSeen := TRUE; END_IF;
        ASSERT_FALSE(fb.RawButton, 'Aucun front pendant bagotement');
ADVANCE_TIME(10000000); fb();
        IF fb.RawX < 5000 THEN oscillationSeen := TRUE; END_IF;
        ASSERT_FALSE(fb.RawButton, 'Aucun front pendant bagotement');
ADVANCE_TIME(10000000); fb();
        IF fb.RawX < 5000 THEN oscillationSeen := TRUE; END_IF;
        ASSERT_FALSE(fb.RawButton, 'Aucun front pendant bagotement');
ADVANCE_TIME(10000000); fb();
        IF fb.RawX < 5000 THEN oscillationSeen := TRUE; END_IF;
        ASSERT_FALSE(fb.RawButton, 'Aucun front pendant bagotement');
ADVANCE_TIME(10000000); fb();
        IF fb.RawX < 5000 THEN oscillationSeen := TRUE; END_IF;
        ASSERT_FALSE(fb.RawButton, 'Aucun front pendant bagotement');
ADVANCE_TIME(10000000); fb();
        IF fb.RawX < 5000 THEN oscillationSeen := TRUE; END_IF;
        ASSERT_FALSE(fb.RawButton, 'Aucun front pendant bagotement');
ADVANCE_TIME(10000000); fb();
        IF fb.RawX < 5000 THEN oscillationSeen := TRUE; END_IF;
        ASSERT_FALSE(fb.RawButton, 'Aucun front pendant bagotement');
ADVANCE_TIME(10000000); fb();
        IF fb.RawX < 5000 THEN oscillationSeen := TRUE; END_IF;
        ASSERT_FALSE(fb.RawButton, 'Aucun front pendant bagotement');
ADVANCE_TIME(10000000); fb();
        IF fb.RawX < 5000 THEN oscillationSeen := TRUE; END_IF;
        ASSERT_FALSE(fb.RawButton, 'Aucun front pendant bagotement');
ADVANCE_TIME(10000000); fb();
        IF fb.RawX < 5000 THEN oscillationSeen := TRUE; END_IF;
        ASSERT_FALSE(fb.RawButton, 'Aucun front pendant bagotement');
ADVANCE_TIME(10000000); fb();
        IF fb.RawX < 5000 THEN oscillationSeen := TRUE; END_IF;
        ASSERT_FALSE(fb.RawButton, 'Aucun front pendant bagotement');
ADVANCE_TIME(10000000); fb();
        IF fb.RawX < 5000 THEN oscillationSeen := TRUE; END_IF;
        ASSERT_FALSE(fb.RawButton, 'Aucun front pendant bagotement');
ADVANCE_TIME(10000000); fb();
        IF fb.RawX < 5000 THEN oscillationSeen := TRUE; END_IF;
        ASSERT_FALSE(fb.RawButton, 'Aucun front pendant bagotement');
ADVANCE_TIME(10000000); fb();
        IF fb.RawX < 5000 THEN oscillationSeen := TRUE; END_IF;
        ASSERT_FALSE(fb.RawButton, 'Aucun front pendant bagotement');
ADVANCE_TIME(10000000); fb();
        IF fb.RawX < 5000 THEN oscillationSeen := TRUE; END_IF;
        ASSERT_FALSE(fb.RawButton, 'Aucun front pendant bagotement');
ADVANCE_TIME(10000000); fb();
        IF fb.RawX < 5000 THEN oscillationSeen := TRUE; END_IF;
        ASSERT_FALSE(fb.RawButton, 'Aucun front pendant bagotement');
ADVANCE_TIME(10000000); fb();
        IF fb.RawX < 5000 THEN oscillationSeen := TRUE; END_IF;
        ASSERT_FALSE(fb.RawButton, 'Aucun front pendant bagotement');
ADVANCE_TIME(10000000); fb();
        IF fb.RawX < 5000 THEN oscillationSeen := TRUE; END_IF;
        ASSERT_FALSE(fb.RawButton, 'Aucun front pendant bagotement');
ADVANCE_TIME(10000000); fb();
        IF fb.RawX < 5000 THEN oscillationSeen := TRUE; END_IF;
        ASSERT_FALSE(fb.RawButton, 'Aucun front pendant bagotement');
ADVANCE_TIME(10000000); fb();
        IF fb.RawX < 5000 THEN oscillationSeen := TRUE; END_IF;
        ASSERT_FALSE(fb.RawButton, 'Aucun front pendant bagotement');
ADVANCE_TIME(10000000); fb();
        IF fb.RawX < 5000 THEN oscillationSeen := TRUE; END_IF;
        ASSERT_FALSE(fb.RawButton, 'Aucun front pendant bagotement');
ADVANCE_TIME(10000000); fb();
        IF fb.RawX < 5000 THEN oscillationSeen := TRUE; END_IF;
        ASSERT_FALSE(fb.RawButton, 'Aucun front pendant bagotement');
ADVANCE_TIME(10000000); fb();
        IF fb.RawX < 5000 THEN oscillationSeen := TRUE; END_IF;
        ASSERT_FALSE(fb.RawButton, 'Aucun front pendant bagotement');
ADVANCE_TIME(10000000); fb();
        IF fb.RawX < 5000 THEN oscillationSeen := TRUE; END_IF;
        ASSERT_FALSE(fb.RawButton, 'Aucun front pendant bagotement');
ADVANCE_TIME(10000000); fb();
        IF fb.RawX < 5000 THEN oscillationSeen := TRUE; END_IF;
        ASSERT_FALSE(fb.RawButton, 'Aucun front pendant bagotement');
ADVANCE_TIME(10000000); fb();
        IF fb.RawX < 5000 THEN oscillationSeen := TRUE; END_IF;
        ASSERT_FALSE(fb.RawButton, 'Aucun front pendant bagotement');
ADVANCE_TIME(10000000); fb();
        IF fb.RawX < 5000 THEN oscillationSeen := TRUE; END_IF;
        ASSERT_FALSE(fb.RawButton, 'Aucun front pendant bagotement');
ADVANCE_TIME(10000000); fb();
        IF fb.RawX < 5000 THEN oscillationSeen := TRUE; END_IF;
        ASSERT_FALSE(fb.RawButton, 'Aucun front pendant bagotement');
ADVANCE_TIME(10000000); fb();
        IF fb.RawX < 5000 THEN oscillationSeen := TRUE; END_IF;
        ASSERT_FALSE(fb.RawButton, 'Aucun front pendant bagotement');
ADVANCE_TIME(10000000); fb();
        IF fb.RawX < 5000 THEN oscillationSeen := TRUE; END_IF;
        ASSERT_FALSE(fb.RawButton, 'Aucun front pendant bagotement');
ADVANCE_TIME(10000000); fb();
        IF fb.RawX < 5000 THEN oscillationSeen := TRUE; END_IF;
        ASSERT_FALSE(fb.RawButton, 'Aucun front pendant bagotement');
ADVANCE_TIME(10000000); fb();
        IF fb.RawX < 5000 THEN oscillationSeen := TRUE; END_IF;
        ASSERT_FALSE(fb.RawButton, 'Aucun front pendant bagotement');
ADVANCE_TIME(10000000); fb();
        IF fb.RawX < 5000 THEN oscillationSeen := TRUE; END_IF;
        ASSERT_FALSE(fb.RawButton, 'Aucun front pendant bagotement');
ADVANCE_TIME(10000000); fb();
        IF fb.RawX < 5000 THEN oscillationSeen := TRUE; END_IF;
        ASSERT_FALSE(fb.RawButton, 'Aucun front pendant bagotement');
ADVANCE_TIME(10000000); fb();
        IF fb.RawX < 5000 THEN oscillationSeen := TRUE; END_IF;
        ASSERT_FALSE(fb.RawButton, 'Aucun front pendant bagotement');
ADVANCE_TIME(10000000); fb();
        IF fb.RawX < 5000 THEN oscillationSeen := TRUE; END_IF;
        ASSERT_FALSE(fb.RawButton, 'Aucun front pendant bagotement');
ADVANCE_TIME(10000000); fb();
        IF fb.RawX < 5000 THEN oscillationSeen := TRUE; END_IF;
        ASSERT_FALSE(fb.RawButton, 'Aucun front pendant bagotement');
ADVANCE_TIME(10000000); fb();
        IF fb.RawX < 5000 THEN oscillationSeen := TRUE; END_IF;
        ASSERT_FALSE(fb.RawButton, 'Aucun front pendant bagotement');
ADVANCE_TIME(10000000); fb();
        IF fb.RawX < 5000 THEN oscillationSeen := TRUE; END_IF;
        ASSERT_FALSE(fb.RawButton, 'Aucun front pendant bagotement');
ADVANCE_TIME(10000000); fb();
        IF fb.RawX < 5000 THEN oscillationSeen := TRUE; END_IF;
        ASSERT_FALSE(fb.RawButton, 'Aucun front pendant bagotement');
ADVANCE_TIME(10000000); fb();
        IF fb.RawX < 5000 THEN oscillationSeen := TRUE; END_IF;
        ASSERT_FALSE(fb.RawButton, 'Aucun front pendant bagotement');
ADVANCE_TIME(10000000); fb();
        IF fb.RawX < 5000 THEN oscillationSeen := TRUE; END_IF;
        ASSERT_FALSE(fb.RawButton, 'Aucun front pendant bagotement');
ADVANCE_TIME(10000000); fb();
        IF fb.RawX < 5000 THEN oscillationSeen := TRUE; END_IF;
        ASSERT_FALSE(fb.RawButton, 'Aucun front pendant bagotement');
ADVANCE_TIME(10000000); fb();
        IF fb.RawX < 5000 THEN oscillationSeen := TRUE; END_IF;
        ASSERT_FALSE(fb.RawButton, 'Aucun front pendant bagotement');
ADVANCE_TIME(10000000); fb();
        IF fb.RawX < 5000 THEN oscillationSeen := TRUE; END_IF;
        ASSERT_FALSE(fb.RawButton, 'Aucun front pendant bagotement');
ADVANCE_TIME(10000000); fb();
        IF fb.RawX < 5000 THEN oscillationSeen := TRUE; END_IF;
        ASSERT_FALSE(fb.RawButton, 'Aucun front pendant bagotement');
ADVANCE_TIME(10000000); fb();
        IF fb.RawX < 5000 THEN oscillationSeen := TRUE; END_IF;
        ASSERT_FALSE(fb.RawButton, 'Aucun front pendant bagotement');
ADVANCE_TIME(10000000); fb();
        IF fb.RawX < 5000 THEN oscillationSeen := TRUE; END_IF;
        ASSERT_FALSE(fb.RawButton, 'Aucun front pendant bagotement');
ADVANCE_TIME(10000000); fb();
        IF fb.RawX < 5000 THEN oscillationSeen := TRUE; END_IF;
        ASSERT_FALSE(fb.RawButton, 'Aucun front pendant bagotement');
ADVANCE_TIME(10000000); fb();
        IF fb.RawX < 5000 THEN oscillationSeen := TRUE; END_IF;
        ASSERT_FALSE(fb.RawButton, 'Aucun front pendant bagotement');
ADVANCE_TIME(10000000); fb();
        IF fb.RawX < 5000 THEN oscillationSeen := TRUE; END_IF;
        ASSERT_FALSE(fb.RawButton, 'Aucun front pendant bagotement');
ADVANCE_TIME(10000000); fb();
        IF fb.RawX < 5000 THEN oscillationSeen := TRUE; END_IF;
        ASSERT_FALSE(fb.RawButton, 'Aucun front pendant bagotement');
ADVANCE_TIME(10000000); fb();
        IF fb.RawX < 5000 THEN oscillationSeen := TRUE; END_IF;
        ASSERT_FALSE(fb.RawButton, 'Aucun front pendant bagotement');
ADVANCE_TIME(10000000); fb();
        IF fb.RawX < 5000 THEN oscillationSeen := TRUE; END_IF;
        ASSERT_FALSE(fb.RawButton, 'Aucun front pendant bagotement');
ADVANCE_TIME(10000000); fb();
        IF fb.RawX < 5000 THEN oscillationSeen := TRUE; END_IF;
        ASSERT_FALSE(fb.RawButton, 'Aucun front pendant bagotement');
ADVANCE_TIME(10000000); fb();
        IF fb.RawX < 5000 THEN oscillationSeen := TRUE; END_IF;
        ASSERT_FALSE(fb.RawButton, 'Aucun front pendant bagotement');
ADVANCE_TIME(10000000); fb();
        IF fb.RawX < 5000 THEN oscillationSeen := TRUE; END_IF;
        ASSERT_FALSE(fb.RawButton, 'Aucun front pendant bagotement');
ADVANCE_TIME(10000000); fb();
        IF fb.RawX < 5000 THEN oscillationSeen := TRUE; END_IF;
        ASSERT_FALSE(fb.RawButton, 'Aucun front pendant bagotement');
ADVANCE_TIME(10000000); fb();
        IF fb.RawX < 5000 THEN oscillationSeen := TRUE; END_IF;
        ASSERT_FALSE(fb.RawButton, 'Aucun front pendant bagotement');
ADVANCE_TIME(10000000); fb();
        IF fb.RawX < 5000 THEN oscillationSeen := TRUE; END_IF;
        ASSERT_FALSE(fb.RawButton, 'Aucun front pendant bagotement');
ADVANCE_TIME(10000000); fb();
        IF fb.RawX < 5000 THEN oscillationSeen := TRUE; END_IF;
        ASSERT_FALSE(fb.RawButton, 'Aucun front pendant bagotement');
ADVANCE_TIME(10000000); fb();
        IF fb.RawX < 5000 THEN oscillationSeen := TRUE; END_IF;
        ASSERT_FALSE(fb.RawButton, 'Aucun front pendant bagotement');
ADVANCE_TIME(10000000); fb();
        IF fb.RawX < 5000 THEN oscillationSeen := TRUE; END_IF;
        ASSERT_FALSE(fb.RawButton, 'Aucun front pendant bagotement');
ADVANCE_TIME(10000000); fb();
        IF fb.RawX < 5000 THEN oscillationSeen := TRUE; END_IF;
        ASSERT_FALSE(fb.RawButton, 'Aucun front pendant bagotement');
ADVANCE_TIME(10000000); fb();
        IF fb.RawX < 5000 THEN oscillationSeen := TRUE; END_IF;
        ASSERT_FALSE(fb.RawButton, 'Aucun front pendant bagotement');
ADVANCE_TIME(10000000); fb();
        IF fb.RawX < 5000 THEN oscillationSeen := TRUE; END_IF;
        ASSERT_FALSE(fb.RawButton, 'Aucun front pendant bagotement');
ADVANCE_TIME(10000000); fb();
        IF fb.RawX < 5000 THEN oscillationSeen := TRUE; END_IF;
        ASSERT_FALSE(fb.RawButton, 'Aucun front pendant bagotement');
ADVANCE_TIME(10000000); fb();
        IF fb.RawX < 5000 THEN oscillationSeen := TRUE; END_IF;
        ASSERT_FALSE(fb.RawButton, 'Aucun front pendant bagotement');
ADVANCE_TIME(10000000); fb();
        IF fb.RawX < 5000 THEN oscillationSeen := TRUE; END_IF;
        ASSERT_FALSE(fb.RawButton, 'Aucun front pendant bagotement');
ADVANCE_TIME(10000000); fb();
        IF fb.RawX < 5000 THEN oscillationSeen := TRUE; END_IF;
        ASSERT_FALSE(fb.RawButton, 'Aucun front pendant bagotement');
ADVANCE_TIME(10000000); fb();
        IF fb.RawX < 5000 THEN oscillationSeen := TRUE; END_IF;
        ASSERT_FALSE(fb.RawButton, 'Aucun front pendant bagotement');
ADVANCE_TIME(10000000); fb();
        IF fb.RawX < 5000 THEN oscillationSeen := TRUE; END_IF;
        ASSERT_FALSE(fb.RawButton, 'Aucun front pendant bagotement');
ADVANCE_TIME(10000000); fb();
        IF fb.RawX < 5000 THEN oscillationSeen := TRUE; END_IF;
        ASSERT_FALSE(fb.RawButton, 'Aucun front pendant bagotement');
ADVANCE_TIME(10000000); fb();
        IF fb.RawX < 5000 THEN oscillationSeen := TRUE; END_IF;
        ASSERT_FALSE(fb.RawButton, 'Aucun front pendant bagotement');
ADVANCE_TIME(10000000); fb();
        IF fb.RawX < 5000 THEN oscillationSeen := TRUE; END_IF;
        ASSERT_FALSE(fb.RawButton, 'Aucun front pendant bagotement');
ADVANCE_TIME(10000000); fb();
        IF fb.RawX < 5000 THEN oscillationSeen := TRUE; END_IF;
        ASSERT_FALSE(fb.RawButton, 'Aucun front pendant bagotement');
ADVANCE_TIME(10000000); fb();
        IF fb.RawX < 5000 THEN oscillationSeen := TRUE; END_IF;
        ASSERT_FALSE(fb.RawButton, 'Aucun front pendant bagotement');
ADVANCE_TIME(10000000); fb();
        IF fb.RawX < 5000 THEN oscillationSeen := TRUE; END_IF;
        ASSERT_FALSE(fb.RawButton, 'Aucun front pendant bagotement');
ADVANCE_TIME(10000000); fb();
        IF fb.RawX < 5000 THEN oscillationSeen := TRUE; END_IF;
        ASSERT_FALSE(fb.RawButton, 'Aucun front pendant bagotement');
ADVANCE_TIME(10000000); fb();
        IF fb.RawX < 5000 THEN oscillationSeen := TRUE; END_IF;
        ASSERT_FALSE(fb.RawButton, 'Aucun front pendant bagotement');
ADVANCE_TIME(10000000); fb();
        IF fb.RawX < 5000 THEN oscillationSeen := TRUE; END_IF;
        ASSERT_FALSE(fb.RawButton, 'Aucun front pendant bagotement');
ADVANCE_TIME(10000000); fb();
        IF fb.RawX < 5000 THEN oscillationSeen := TRUE; END_IF;
        ASSERT_FALSE(fb.RawButton, 'Aucun front pendant bagotement');
ADVANCE_TIME(10000000); fb();
        IF fb.RawX < 5000 THEN oscillationSeen := TRUE; END_IF;
        ASSERT_FALSE(fb.RawButton, 'Aucun front pendant bagotement');
ADVANCE_TIME(10000000); fb();
        IF fb.RawX < 5000 THEN oscillationSeen := TRUE; END_IF;
        ASSERT_FALSE(fb.RawButton, 'Aucun front pendant bagotement');
ADVANCE_TIME(10000000); fb();
        IF fb.RawX < 5000 THEN oscillationSeen := TRUE; END_IF;
        ASSERT_FALSE(fb.RawButton, 'Aucun front pendant bagotement');
ADVANCE_TIME(10000000); fb();
        IF fb.RawX < 5000 THEN oscillationSeen := TRUE; END_IF;
        ASSERT_FALSE(fb.RawButton, 'Aucun front pendant bagotement');
ADVANCE_TIME(10000000); fb();
        IF fb.RawX < 5000 THEN oscillationSeen := TRUE; END_IF;
        ASSERT_FALSE(fb.RawButton, 'Aucun front pendant bagotement');
ADVANCE_TIME(10000000); fb();
        IF fb.RawX < 5000 THEN oscillationSeen := TRUE; END_IF;
        ASSERT_FALSE(fb.RawButton, 'Aucun front pendant bagotement');
ADVANCE_TIME(10000000); fb();
        IF fb.RawX < 5000 THEN oscillationSeen := TRUE; END_IF;
        ASSERT_FALSE(fb.RawButton, 'Aucun front pendant bagotement');
ADVANCE_TIME(10000000); fb();
        IF fb.RawX < 5000 THEN oscillationSeen := TRUE; END_IF;
        ASSERT_FALSE(fb.RawButton, 'Aucun front pendant bagotement');
ADVANCE_TIME(10000000); fb();
        IF fb.RawX < 5000 THEN oscillationSeen := TRUE; END_IF;
        ASSERT_FALSE(fb.RawButton, 'Aucun front pendant bagotement');
ADVANCE_TIME(10000000); fb();
        IF fb.RawX < 5000 THEN oscillationSeen := TRUE; END_IF;
        ASSERT_FALSE(fb.RawButton, 'Aucun front pendant bagotement');
ADVANCE_TIME(10000000); fb();
        IF fb.RawX < 5000 THEN oscillationSeen := TRUE; END_IF;
        ASSERT_FALSE(fb.RawButton, 'Aucun front pendant bagotement');
ADVANCE_TIME(10000000); fb();
        IF fb.RawX < 5000 THEN oscillationSeen := TRUE; END_IF;
        ASSERT_FALSE(fb.RawButton, 'Aucun front pendant bagotement');
ADVANCE_TIME(10000000); fb();
        IF fb.RawX < 5000 THEN oscillationSeen := TRUE; END_IF;
        ASSERT_FALSE(fb.RawButton, 'Aucun front pendant bagotement');
ADVANCE_TIME(10000000); fb();
        IF fb.RawX < 5000 THEN oscillationSeen := TRUE; END_IF;
        ASSERT_FALSE(fb.RawButton, 'Aucun front pendant bagotement');
ADVANCE_TIME(10000000); fb();
        IF fb.RawX < 5000 THEN oscillationSeen := TRUE; END_IF;
        ASSERT_FALSE(fb.RawButton, 'Aucun front pendant bagotement');
ADVANCE_TIME(10000000); fb();
        IF fb.RawX < 5000 THEN oscillationSeen := TRUE; END_IF;
        ASSERT_FALSE(fb.RawButton, 'Aucun front pendant bagotement');
ADVANCE_TIME(10000000); fb();
        IF fb.RawX < 5000 THEN oscillationSeen := TRUE; END_IF;
        ASSERT_FALSE(fb.RawButton, 'Aucun front pendant bagotement');
ADVANCE_TIME(10000000); fb();
        IF fb.RawX < 5000 THEN oscillationSeen := TRUE; END_IF;
        ASSERT_FALSE(fb.RawButton, 'Aucun front pendant bagotement');
ADVANCE_TIME(10000000); fb();
        IF fb.RawX < 5000 THEN oscillationSeen := TRUE; END_IF;
        ASSERT_FALSE(fb.RawButton, 'Aucun front pendant bagotement');
ADVANCE_TIME(10000000); fb();
        IF fb.RawX < 5000 THEN oscillationSeen := TRUE; END_IF;
        ASSERT_FALSE(fb.RawButton, 'Aucun front pendant bagotement');
ADVANCE_TIME(10000000); fb();
        IF fb.RawX < 5000 THEN oscillationSeen := TRUE; END_IF;
        ASSERT_FALSE(fb.RawButton, 'Aucun front pendant bagotement');
ADVANCE_TIME(10000000); fb();
        IF fb.RawX < 5000 THEN oscillationSeen := TRUE; END_IF;
        ASSERT_FALSE(fb.RawButton, 'Aucun front pendant bagotement');
ADVANCE_TIME(10000000); fb();
        IF fb.RawX < 5000 THEN oscillationSeen := TRUE; END_IF;
        ASSERT_FALSE(fb.RawButton, 'Aucun front pendant bagotement');
ADVANCE_TIME(10000000); fb();
        IF fb.RawX < 5000 THEN oscillationSeen := TRUE; END_IF;
        ASSERT_FALSE(fb.RawButton, 'Aucun front pendant bagotement');
ADVANCE_TIME(10000000); fb();
        IF fb.RawX < 5000 THEN oscillationSeen := TRUE; END_IF;
        ASSERT_FALSE(fb.RawButton, 'Aucun front pendant bagotement');
ADVANCE_TIME(10000000); fb();
        IF fb.RawX < 5000 THEN oscillationSeen := TRUE; END_IF;
        ASSERT_FALSE(fb.RawButton, 'Aucun front pendant bagotement');
ADVANCE_TIME(10000000); fb();
        IF fb.RawX < 5000 THEN oscillationSeen := TRUE; END_IF;
        ASSERT_FALSE(fb.RawButton, 'Aucun front pendant bagotement');
ADVANCE_TIME(10000000); fb();
        IF fb.RawX < 5000 THEN oscillationSeen := TRUE; END_IF;
        ASSERT_FALSE(fb.RawButton, 'Aucun front pendant bagotement');
ADVANCE_TIME(10000000); fb();
        IF fb.RawX < 5000 THEN oscillationSeen := TRUE; END_IF;
        ASSERT_FALSE(fb.RawButton, 'Aucun front pendant bagotement');
ADVANCE_TIME(10000000); fb();
        IF fb.RawX < 5000 THEN oscillationSeen := TRUE; END_IF;
        ASSERT_FALSE(fb.RawButton, 'Aucun front pendant bagotement');
ADVANCE_TIME(10000000); fb();
        IF fb.RawX < 5000 THEN oscillationSeen := TRUE; END_IF;
        ASSERT_FALSE(fb.RawButton, 'Aucun front pendant bagotement');
ADVANCE_TIME(10000000); fb();
        IF fb.RawX < 5000 THEN oscillationSeen := TRUE; END_IF;
        ASSERT_FALSE(fb.RawButton, 'Aucun front pendant bagotement');
ADVANCE_TIME(10000000); fb();
        IF fb.RawX < 5000 THEN oscillationSeen := TRUE; END_IF;
        ASSERT_FALSE(fb.RawButton, 'Aucun front pendant bagotement');
ADVANCE_TIME(10000000); fb();
        IF fb.RawX < 5000 THEN oscillationSeen := TRUE; END_IF;
        ASSERT_FALSE(fb.RawButton, 'Aucun front pendant bagotement');
ADVANCE_TIME(10000000); fb();
        IF fb.RawX < 5000 THEN oscillationSeen := TRUE; END_IF;
        ASSERT_FALSE(fb.RawButton, 'Aucun front pendant bagotement');
ADVANCE_TIME(10000000); fb();
        IF fb.RawX < 5000 THEN oscillationSeen := TRUE; END_IF;
        ASSERT_FALSE(fb.RawButton, 'Aucun front pendant bagotement');
ADVANCE_TIME(10000000); fb();
        IF fb.RawX < 5000 THEN oscillationSeen := TRUE; END_IF;
        ASSERT_FALSE(fb.RawButton, 'Aucun front pendant bagotement');
ADVANCE_TIME(10000000); fb();
        IF fb.RawX < 5000 THEN oscillationSeen := TRUE; END_IF;
        ASSERT_FALSE(fb.RawButton, 'Aucun front pendant bagotement');
ADVANCE_TIME(10000000); fb();
        IF fb.RawX < 5000 THEN oscillationSeen := TRUE; END_IF;
        ASSERT_FALSE(fb.RawButton, 'Aucun front pendant bagotement');
    ASSERT_TRUE(oscillationSeen, 'Bagotement traverse le neutre');
    ASSERT_EQ(fb.RawX, 5000, 'Bagotement stabilise');
END_TEST
